  end
  visorFuncEasyPick_b634ba()
  # end: URCap Program Node
  $ 1699 "MoveJ"
  $ 1700 "Waypoint_95" "breakAfter"
  movej(get_inverse_kin(Waypoint_95_p, qnear=Waypoint_95_q), a=1.3962634015954636, v=1.0471975511965976)
  $ 1701 "Wait: 2.0"
  sleep(2.0)
  elif (7 == switch_1):
    $ 1702 "Case 7"
  elif (8 == switch_1):
    $ 1731 "Case 8"
  elif (11 == switch_1):
    $ 1764 "Case 11"
  elif (12 == switch_1):
    $ 1801 "Case 12"
  elif (15 == switch_1):
    $ 1852 "Case 15"
  elif (30 == switch_1):
    $ 1855 "Case 30"
  elif (31 == switch_1):
    $ 1888 "Case 31"
  elif (32 == switch_1):
    $ 1900 "Case 32"
  elif (33 == switch_1):
    $ 1941 "Case 33"
  elif (35 == switch_1):
    $ 2007 "Case 35"
    $ 2008 "Pick the powder container"
    # begin: URCap Program Node
    #   Source: SensoPart VISOR Robotic, 2.0.0, SensoPart Industriesensorik GmbH
    #   Type: VISOR Robotic App
    $ 2011 "VISOR Easy Pick"
    def visorFuncEasyPick_ceefd3():
      # begin: URCap Program Node
      #   Source: SensoPart VISOR Robotic, 2.0.0, SensoPart Industriesensorik GmbH
      #   Type: Easy Pick Setup
      $ 2012 "# 1 Setup" "noBreak"
      local easyPickVisorId = 1
      local easyPickArmMounted = True
      local easyPickSetJob = True
      local easyPickJobName = "Container"
      local easyPickAtImgAcq = False
      local easyPickImgAcqPose = cont_img_pose
      # end: URCap Program Node
      # begin: URCap Program Node
      #   Source: SensoPart VISOR Robotic, 2.0.0, SensoPart Industriesensorik GmbH
      #   Type: Process
      $ 2013 "Process" "noBreak"
      local easyPickObjTaken = False
      local easyPickTrigger = False
      local easyPickPoseIdx = 0
      local easyPickPose = p[0,0,0,0,0,0]
      def easyPickFuncTrigger(visorId, setJob, jobName, arm):
      if (setJob):
        visor_changeJob(visorId, jobName, 6000)
      end
      if (arm):
        visor_trigger(visorId, 6000, "arm")
      else:
        visor_trigger(visorId, 6000)
      end
      global easyPickParts=visor_partsFound(visorId)
      visor_easyPickUpdate(visorId, "parts", visor_partsFound(visorId))
      return visor_getPose3d(visorId, 0)
    end
    while (not easyPickObjTaken):
      easyPickTrigger = (easyPickCount >= visor_partsFound(easyPickVisorId)) or (easyPickCount > 9) or (not visor_easyPickCheckIdent("bb1e48", easyPickVisorId))
      if (easyPickTrigger):
        easyPickCount = 0
      end
      easyPickPoseIdx = easyPickCount
      easyPickPose = visor_getPose3d(easyPickVisorId, easyPickPoseIdx)
      visor_easyPickUpdate(easyPickVisorId, "counter", easyPickPoseIdx)
      # begin: URCap Program Node
      #   Source: SensoPart VISOR Robotic, 2.0.0, SensoPart Industriesensorik GmbH
      #   Type: Image Acquisition Pose
      $ 2014 "Image Acquisition Pose" "noBreak"
      if (easyPickTrigger):
        if (not easyPickAtImgAcq):
          movej(pose_trans(easyPickImgAcqPose,p[0.0000,0.0000,-0.0000,0.0000,0.0000,0.0000]),a=1.3963,v=1.0472,t=0.000000,r=0.000000)
          easyPickAtImgAcq = True
        end
        easyPickPose = easyPickFuncTrigger(easyPickVisorId, easyPickSetJob, easyPickJobName, easyPickArmMounted)
      end
      # end: URCap Program Node
      # begin: URCap Program Node
      #   Source: SensoPart VISOR Robotic, 2.0.0, SensoPart Industriesensorik GmbH
      #   Type: Object Detected
      $ 2015 "Object Detected" "noBreak"
      if (visor_partsFound(easyPickVisorId) > 0):
        $ 2016 "Open Gripper" "noBreak"
        # begin: URCap Program Node
        #   Source: Robotiq_Grippers, 1.8.4.4844, Robotiq Inc.
        #   Type: Gripper
        $ 2017 "Gripper Open (1)" "noBreak"
        if not(gripper_connected[0]):
          popup("Gripper 1 must be connected to run this program.", "No connection", False, True, True)
        end
        if not(rq_is_gripper_activated("1")):
          popup("Gripper 1 is not activated. Go to Installation tab > Gripper to activate it and run the program again.", "Not activated", False, True, True)
        end
        rq_set_pos_spd_for(0, 102, 77, "1")
        rq_wait_pos_spe_for_request(0, 102, 77, "1")
        rq_go_to("1")
        rq_wait("1")
        # end: URCap Program Node
        $ 2018 "MoveJ" "noBreak"
        $ 2019 "Waypoint_13" "noBreak"
        movej(get_inverse_kin(Waypoint_13_p, qnear=Waypoint_13_q), a=1.3962634015954636, v=1.0471975511965976)
        # begin: URCap Program Node
        #   Source: SensoPart VISOR Robotic, 2.0.0, SensoPart Industriesensorik GmbH
        #   Type: Approach Pose
        $ 2020 "Approach Pose" "noBreak"
        movej(pose_trans(easyPickPose,p[0.0000,0.0000,0.0500,0.0000,0.0000,0.0000]),a=1.3963,v=1.0472,t=0.000000,r=0.000000)
        # end: URCap Program Node
        # begin: URCap Program Node
        #   Source: SensoPart VISOR Robotic, 2.0.0, SensoPart Industriesensorik GmbH
        #   Type: Target Pose
        $ 2021 "Target Pose" "noBreak"
        movel(pose_trans(easyPickPose,p[0.0000,0.0000,-0.0000,0.0000,0.0000,0.0000]),a=0.5000,v=0.2500,t=0.000000,r=0.000000)
        # end: URCap Program Node
        $ 2022 "Close Gripper" "noBreak"
        # begin: URCap Program Node
        #   Source: Robotiq_Grippers, 1.8.4.4844, Robotiq Inc.
        #   Type: Gripper
        $ 2023 "Gripper Close (1)" "noBreak"
        if not(gripper_connected[0]):
          popup("Gripper 1 must be connected to run this program.", "No connection", False, True, True)
        end
        if not(rq_is_gripper_activated("1")):
          popup("Gripper 1 is not activated. Go to Installation tab > Gripper to activate it and run the program again.", "Not activated", False, True, True)
        end
        rq_set_pos_spd_for(255, 102, 77, "1")
        rq_wait_pos_spe_for_request(255, 102, 77, "1")
        rq_go_to("1")
        rq_wait("1")
        # end: URCap Program Node
        # begin: URCap Program Node
        #   Source: SensoPart VISOR Robotic, 2.0.0, SensoPart Industriesensorik GmbH
        #   Type: Exit Pose
        $ 2024 "Exit Pose" "noBreak"
        movel(pose_trans(easyPickPose,p[0.0000,0.0000,0.0500,0.0000,0.0000,0.0000]),a=0.5000,v=0.2500,t=0.000000,r=0.000000)
        # end: URCap Program Node
        easyPickObjTaken = True
      end
      # end: URCap Program Node
      # begin: URCap Program Node
      #   Source: SensoPart VISOR Robotic, 2.0.0, SensoPart Industriesensorik GmbH
      #   Type: No Object Detected
      $ 2025 "No Object Detected" "noBreak"
      if (visor_partsFound(easyPickVisorId) < 1):
        $ 2026 "Popup: No Container detected" "noBreak"
        popup("No Container detected", "Message", False, False, blocking=True)
        else:
      end
      # end: URCap Program Node
    end
    easyPickCount = easyPickCount + 1
    visor_easyPickUpdate(easyPickVisorId, "counter", easyPickCount)
    visor_easyPickSetIdent("bb1e48", easyPickVisorId)
    # end: URCap Program Node
  end
  visorFuncEasyPick_ceefd3()
  # end: URCap Program Node
  $ 2027 "MoveJ"
  $ 2029 "Waypoint_70" "breakAfter"
  movej(get_inverse_kin(Waypoint_70_p, qnear=Waypoint_70_q), a=0.6981317007977318, v=0.5235987755982988)
  $ 2030 "Waypoint_2" "breakAfter"
  movej(get_inverse_kin(Waypoint_2_p, qnear=Waypoint_2_q), a=0.8726646259971648, v=0.5235987755982988, r=0.05)
  $ 2031 "Waypoint_3" "breakAfter"
  movej(get_inverse_kin(Waypoint_3_p, qnear=Waypoint_3_q), a=0.6981317007977318, v=0.5235987755982988, r=0.05)
  $ 2032 "MoveL"
  $ 2033 "Waypoint_15" "breakAfter"
  movel(Waypoint_15_p, a=0.5, v=0.1, r=0.05)
  $ 2034 "Waypoint_14" "breakAfter"
  movel(Waypoint_14_p, a=0.3, v=0.1)
  $ 2035 "Waypoint_4" "breakAfter"
  movel(Waypoint_4_p, a=0.3, v=0.05)
  # begin: URCap Program Node
  #   Source: Robotiq_Grippers, 1.8.4.4844, Robotiq Inc.
  #   Type: Gripper
  $ 2036 "Gripper Open (1)"
  if not(gripper_connected[0]):
    popup("Gripper 1 must be connected to run this program.", "No connection", False, True, True)
  end
  if not(rq_is_gripper_activated("1")):
    popup("Gripper 1 is not activated. Go to Installation tab > Gripper to activate it and run the program again.", "Not activated", False, True, True)
  end
  rq_set_pos_spd_for(0, 102, 77, "1")
  rq_wait_pos_spe_for_request(0, 102, 77, "1")
  rq_go_to("1")
  rq_wait("1")
  # end: URCap Program Node
  $ 2037 "MoveL"
  $ 2038 "Waypoint_25" "breakAfter"
  movel(Waypoint_25_p, a=0.3, v=0.1)
  $ 2039 "Waypoint_15" "breakAfter"
  movel(Waypoint_15_p, a=0.5, v=0.1, r=0.05)
  $ 2040 "Home (Safe)"
  movej([-1.2302089344500047, -1.2969853503591224, -1.875639182904262, -1.539621866126728, 1.5731943360401213, -2.80099559440227], a=1.3962634015954636, v=1.0471975511965976)
  elif (36 == switch_1):
    $ 2070 "Case 36"
    $ 2074 "Decap"
    $ 2112 "MoveJ"
    $ 2113 "Waypoint_39" "breakAfter"
    movej(get_inverse_kin(Waypoint_39_p, qnear=Waypoint_39_q), a=1.3962634015954636, v=1.0471975511965976)
    $ 2114 "MoveL"
    $ 2115 "Waypoint_41" "breakAfter"
    movel(Waypoint_41_p, a=0.5, v=0.1)
    $ 2116 "Waypoint_40" "breakAfter"
    movel(Waypoint_40_p, a=0.3, v=0.05)
    # begin: URCap Program Node
    #   Source: Robotiq_Grippers, 1.8.4.4844, Robotiq Inc.
    #   Type: Gripper
    $ 2117 "Gripper Close (1)"
    if not(gripper_connected[0]):
      popup("Gripper 1 must be connected to run this program.", "No connection", False, True, True)
    end
    if not(rq_is_gripper_activated("1")):
      popup("Gripper 1 is not activated. Go to Installation tab > Gripper to activate it and run the program again.", "Not activated", False, True, True)
    end
    rq_set_pos_spd_for(255, 77, 51, "1")
    rq_wait_pos_spe_for_request(255, 77, 51, "1")
    rq_go_to("1")
    rq_wait("1")
    # end: URCap Program Node
    $ 2118 "Loop 2 times"
    Loop_2 = 0
    while (Loop_2 < 2):
      $ 2119 "MoveL"
      $ 2120 "Waypoint_42" "breakAfter"
      movel(Waypoint_42_p, a=1.2, v=0.5)
      $ 2121 "Waypoint_43" "breakAfter"
      movel(Waypoint_43_p, a=1.2, v=0.25)
      # begin: URCap Program Node
      #   Source: Robotiq_Grippers, 1.8.4.4844, Robotiq Inc.
      #   Type: Gripper
      $ 2122 "Gripper Move40mm (1)"
      if not(gripper_connected[0]):
        popup("Gripper 1 must be connected to run this program.", "No connection", False, True, True)
      end
      if not(rq_is_gripper_activated("1")):
        popup("Gripper 1 is not activated. Go to Installation tab > Gripper to activate it and run the program again.", "Not activated", False, True, True)
      end
      rq_set_pos_spd_for(63, 77, 51, "1")
      rq_wait_pos_spe_for_request(63, 77, 51, "1")
      rq_go_to("1")
      rq_wait("1")
      # end: URCap Program Node
      $ 2123 "MoveL"
      $ 2124 "Waypoint_44" "breakAfter"
      movel(Waypoint_44_p, a=1.2, v=0.5)
      $ 2125 "Waypoint_45" "breakAfter"
      movel(Waypoint_45_p, a=1.2, v=0.25)
      # begin: URCap Program Node
      #   Source: Robotiq_Grippers, 1.8.4.4844, Robotiq Inc.
      #   Type: Gripper
      $ 2126 "Gripper Move11mm (1)"
      if not(gripper_connected[0]):
        popup("Gripper 1 must be connected to run this program.", "No connection", False, True, True)
      end
      if not(rq_is_gripper_activated("1")):
        popup("Gripper 1 is not activated. Go to Installation tab > Gripper to activate it and run the program again.", "Not activated", False, True, True)
      end
      rq_set_pos_spd_for(200, 77, 51, "1")
      rq_wait_pos_spe_for_request(200, 77, 51, "1")
      rq_go_to("1")
      rq_wait("1")
      # end: URCap Program Node
      Loop_2 = Loop_2 + 1
    end
    $ 2127 "MoveL"
    $ 2128 "Waypoint_46" "breakAfter"
    movel(Waypoint_46_p, a=0.3, v=0.05)
    $ 2129 "Waypoint_47" "breakAfter"
    movel(Waypoint_47_p, a=0.5, v=0.1)
    $ 2130 "Waypoint_48" "breakAfter"
    movel(Waypoint_48_p, a=1.2, v=0.25)
    $ 2131 "Waypoint_49" "breakAfter"
    movel(Waypoint_49_p, a=1.2, v=0.25)
    # begin: URCap Program Node
    #   Source: Robotiq_Grippers, 1.8.4.4844, Robotiq Inc.
    #   Type: Gripper
    $ 2132 "Gripper Move35mm (1)"
    if not(gripper_connected[0]):
      popup("Gripper 1 must be connected to run this program.", "No connection", False, True, True)
    end
    if not(rq_is_gripper_activated("1")):
      popup("Gripper 1 is not activated. Go to Installation tab > Gripper to activate it and run the program again.", "Not activated", False, True, True)
    end
    rq_set_pos_spd_for(87, 77, 51, "1")
    rq_wait_pos_spe_for_request(87, 77, 51, "1")
    rq_go_to("1")
    rq_wait("1")
    # end: URCap Program Node
    $ 2133 "MoveL"
    $ 2134 "Waypoint_50" "breakAfter"
    movel(Waypoint_50_p, a=1.2, v=0.25)
    $ 2135 "Home (Safe)"
    movej([-1.2302089344500047, -1.2969853503591224, -1.875639182904262, -1.539621866126728, 1.5731943360401213, -2.80099559440227], a=1.3962634015954636, v=1.0471975511965976)
  elif (37 == switch_1):
    $ 2136 "Case 37"
    $ 2137 "Powder dispensing"
    $ 2138 "zero_scale()"
    zero_scale()
    # begin: URCap Program Node
    #   Source: SensoPart VISOR Robotic, 2.0.0, SensoPart Industriesensorik GmbH
    #   Type: VISOR Robotic App
    $ 2139 "VISOR Easy Pick"
    def visorFuncEasyPick_f697d2():
      # begin: URCap Program Node
      #   Source: SensoPart VISOR Robotic, 2.0.0, SensoPart Industriesensorik GmbH
      #   Type: Easy Pick Setup
      $ 2140 "# 1 Setup" "noBreak"
      local easyPickVisorId = 1
      local easyPickArmMounted = True
      local easyPickSetJob = True
      local easyPickJobName = "Weigh_scale"
      local easyPickAtImgAcq = False
      local easyPickImgAcqPose = cont_img_pose
      # end: URCap Program Node
      # begin: URCap Program Node
      #   Source: SensoPart VISOR Robotic, 2.0.0, SensoPart Industriesensorik GmbH
      #   Type: Process
      $ 2141 "Process" "noBreak"
      local easyPickObjTaken = False
      local easyPickTrigger = False
      local easyPickPoseIdx = 0
      local easyPickPose = p[0,0,0,0,0,0]
      def easyPickFuncTrigger(visorId, setJob, jobName, arm):
      if (setJob):
        visor_changeJob(visorId, jobName, 6000)
      end
      if (arm):
        visor_trigger(visorId, 6000, "arm")
      else:
        visor_trigger(visorId, 6000)
      end
      global easyPickParts_4=visor_partsFound(visorId)
      visor_easyPickUpdate(visorId, "parts", visor_partsFound(visorId))
      return visor_getPose3d(visorId, 0)
    end
    while (not easyPickObjTaken):
      easyPickTrigger = (easyPickCount_4 >= visor_partsFound(easyPickVisorId)) or (easyPickCount_4 > 9) or (not visor_easyPickCheckIdent("db3fd8", easyPickVisorId))
      if (easyPickTrigger):
        easyPickCount_4 = 0
      end
      easyPickPoseIdx = easyPickCount_4
      easyPickPose = visor_getPose3d(easyPickVisorId, easyPickPoseIdx)
      visor_easyPickUpdate(easyPickVisorId, "counter", easyPickPoseIdx)
      # begin: URCap Program Node
      #   Source: SensoPart VISOR Robotic, 2.0.0, SensoPart Industriesensorik GmbH
      #   Type: Image Acquisition Pose
      $ 2142 "Image Acquisition Pose" "noBreak"
      if (easyPickTrigger):
        if (not easyPickAtImgAcq):
          movej(pose_trans(easyPickImgAcqPose,p[0.0000,0.0000,-0.0000,0.0000,0.0000,0.0000]),a=1.3963,v=1.0472,t=0.000000,r=0.000000)
          easyPickAtImgAcq = True
        end
        easyPickPose = easyPickFuncTrigger(easyPickVisorId, easyPickSetJob, easyPickJobName, easyPickArmMounted)
      end
      # end: URCap Program Node
      # begin: URCap Program Node
      #   Source: SensoPart VISOR Robotic, 2.0.0, SensoPart Industriesensorik GmbH
      #   Type: Object Detected
      $ 2143 "Object Detected" "noBreak"
      if (visor_partsFound(easyPickVisorId) > 0):
        $ 2144 "Open Gripper" "noBreak"
        $ 2145 "MoveL" "noBreak"
        $ 2146 "Weight_value≔get_weight()" "noBreak"
        global Weight_value=get_weight()
        # begin: URCap Program Node
        #   Source: Robotiq_Grippers, 1.8.4.4844, Robotiq Inc.
        #   Type: Gripper
        $ 2147 "Gripper Open (1)" "noBreak"
        if not(gripper_connected[0]):
          popup("Gripper 1 must be connected to run this program.", "No connection", False, True, True)
        end
        if not(rq_is_gripper_activated("1")):
          popup("Gripper 1 is not activated. Go to Installation tab > Gripper to activate it and run the program again.", "Not activated", False, True, True)
        end
        rq_set_pos_spd_for(0, 77, 77, "1")
        rq_wait_pos_spe_for_request(0, 77, 77, "1")
        rq_go_to("1")
        rq_wait("1")
        # end: URCap Program Node
        $ 2148 "Waypoint_53" "noBreak"
        movel(Waypoint_53_p, a=0.6, v=0.15, r=0.05)
        $ 2149 "Spatula_above" "noBreak"
        movel(Spatula_above_p, a=0.6, v=0.15)
        $ 2150 "Spatula_pick" "noBreak"
        movel(Spatula_pick_p, a=0.6, v=0.15)
        # begin: URCap Program Node
        #   Source: Robotiq_Grippers, 1.8.4.4844, Robotiq Inc.
        #   Type: Gripper
        $ 2151 "Gripper Close (1)" "noBreak"
        if not(gripper_connected[0]):
          popup("Gripper 1 must be connected to run this program.", "No connection", False, True, True)
        end
        if not(rq_is_gripper_activated("1")):
          popup("Gripper 1 is not activated. Go to Installation tab > Gripper to activate it and run the program again.", "Not activated", False, True, True)
        end
        rq_set_pos_spd_for(255, 77, 77, "1")
        rq_wait_pos_spe_for_request(255, 77, 77, "1")
        rq_go_to("1")
        rq_wait("1")
        # end: URCap Program Node
        $ 2152 "Spatula_above" "noBreak"
        movel(Spatula_above_p, a=0.6, v=0.15)
        $ 2153 "Popup: Connect the vibration motor" "noBreak"
        popup("Connect the vibration motor", "Message", False, False, blocking=True)
        $ 2154 "tare_scale()" "noBreak"
        tare_scale()
        $ 2155 "container_start" "noBreak"
        movel(container_start_p, a=0.3, v=0.1)
        $ 2156 "container_wp_1" "noBreak"
        movel(container_wp_1_p, a=0.3, v=0.05)
        $ 2157 "Loop 1 times" "noBreak"
        Loop_9 = 0
        while (Loop_9 < 1):
          $ 2158 "Waypoint_55" "noBreak"
          global move_thread_flag_2158=0
          thread move_thread_2158():
            enter_critical
            move_thread_flag_2158 = 1
            movel(Waypoint_55_p, a=0.5, v=0.07)
            move_thread_flag_2158 = 2
            exit_critical
          end
          move_thread_flag_2158 = 0
          move_thread_han_2158 = run move_thread_2158()
          while (True):
            sleep(1.0E-10)
            if (move_thread_flag_2158 > 1):
              join move_thread_han_2158
              break
            end
            sync()
          end
          $ 2160 "Waypoint_56" "noBreak"
          movel(Waypoint_56_p, a=0.3, v=0.05)
          $ 2161 "Waypoint_74" "noBreak"
          movel(Waypoint_74_p, a=0.6, v=0.15)
          $ 2162 "Set AO[0]=3.0" "noBreak"
          set_standard_analog_out(0, 0.3)
          $ 2163 "Wait: 2.0" "noBreak"
          sleep(2.0)
          $ 2164 "Set AO[0]=0.0" "noBreak"
          set_standard_analog_out(0, 0.0)
          Loop_9 = Loop_9 + 1
        end
        $ 2168 "ftr_scoop2" "noBreak"
        movel(ftr_scoop2_p, a=0.3, v=0.05)
        $ 2169 "aftr_scoo3" "noBreak"
        movel(aftr_scoo3_p, a=0.3, v=0.05)
        $ 2170 "MoveJ" "noBreak"
        $ 2171 "Waypoint_60" "noBreak"
        movej(get_inverse_kin(Waypoint_60_p, qnear=Waypoint_60_q), a=0.5235987755982988, v=0.3490658503988659, r=0.05)
        $ 2172 "Waypoint_61" "noBreak"
        movej(get_inverse_kin(Waypoint_61_p, qnear=Waypoint_61_q), a=0.5235987755982988, v=0.3490658503988659, r=0.05)
        # begin: URCap Program Node
        #   Source: SensoPart VISOR Robotic, 2.0.0, SensoPart Industriesensorik GmbH
        #   Type: Approach Pose
        $ 2173 "Approach Pose" "noBreak"
        movej(pose_trans(easyPickPose,p[0.0000,0.0000,0.0500,0.0000,0.0000,0.0000]),a=0.4363,v=0.3491,t=0.000000,r=0.000000)
        # end: URCap Program Node
        # begin: URCap Program Node
        #   Source: SensoPart VISOR Robotic, 2.0.0, SensoPart Industriesensorik GmbH
        #   Type: Target Pose
        $ 2174 "Target Pose" "noBreak"
        movel(pose_trans(easyPickPose,p[0.0000,0.0000,-0.0000,0.0000,0.0000,0.0000]),a=0.1000,v=0.0500,t=0.000000,r=0.000000)
        # end: URCap Program Node
        $ 2175 "Close Gripper" "noBreak"
        $ 2176 "dispense_pos≔get_actual_tcp_pose()" "noBreak"
        global dispense_pos= get_actual_tcp_pose ()
        $ 2177 "MoveL" "noBreak"
        $ 2178 "Start_thread≔ True " "noBreak"
        global Start_thread=  True
        $ 2179 "vib_mot_thread≔ True " "noBreak"
        global vib_mot_thread=  True
        $ 2180 "tilt_angle≔current_pose[4]" "noBreak"
        global tilt_angle=current_pose[4]
        $ 2181 "Wait: 0.5" "noBreak"
        sleep(0.5)
        $ 2182 "Loop Weight_value≤Target_weight and tilt_angle≤-0.40" "noBreak"
        thread Thread_while_2182():
          while (True):
            $ 2183 "current_error≔Target_weight-Weight_value" "noBreak"
            global current_error=Target_weight-Weight_value
            $ 2184 "Integral_error≔Integral_error+current_error*dt" "noBreak"
            global Integral_error=Integral_error+current_error*dt
            $ 2185 "derivative≔(current_error-previous_error)/dt" "noBreak"
            global derivative=(current_error-previous_error)/dt
            $ 2186 "tilt_increment≔(kp*current_error)+(ki*Integral_error)+(kd*derivative)" "noBreak"
            global tilt_increment=(kp*current_error)+(ki*Integral_error)+(kd*derivative)
            $ 2187 "current_pose≔get_actual_tcp_pose()" "noBreak"
            global current_pose= get_actual_tcp_pose ()
            $ 2188 "tilt_angle≔current_pose[4]" "noBreak"
            global tilt_angle=current_pose[4]
            $ 2189 "tilt_pose≔pose_trans(current_pose, p[(tilt_increment/7), 0, 0, 0, tilt_increment, 0])" "noBreak"
            global tilt_pose=pose_trans(current_pose, p[(tilt_increment/7), 0, 0, 0, tilt_increment, 0])
            $ 2190 "movel(tilt_pose, a=0.025, v=0.015, r=0.00001)" "noBreak"
            movel(tilt_pose, a=0.025, v=0.015, r=0.00001)
            $ 2191 "previous_error≔current_error" "noBreak"
            global previous_error=current_error
          end
        end
        if (Weight_value <= Target_weight  and  tilt_angle <= -0.40):
          global thread_handler_2182=run Thread_while_2182()
          while (Weight_value <= Target_weight  and  tilt_angle <= -0.40):
            sync()
          end
          kill thread_handler_2182
        end
        $ 2192 "Start_thread≔ False " "noBreak"
        global Start_thread=  False
        $ 2194 "Weight_value≔get_weight()" "noBreak"
        global Weight_value=get_weight()
        $ 2195 "tilt_angle≔-1" "noBreak"
        global tilt_angle=-1
        $ 2196 "Wait: 0.5" "noBreak"
        sleep(0.5)
        $ 2197 "vib_mot_thread≔ False " "noBreak"
        global vib_mot_thread=  False
        $ 2198 "MoveL" "noBreak"
        $ 2199 "dispense_pos" "noBreak"
        movel(dispense_pos, a=0.2, v=0.05)
        $ 2200 "Integral_error≔0" "noBreak"
        global Integral_error=0
        $ 2201 "current_error≔0" "noBreak"
        global current_error=0
        $ 2202 "previous_error≔0" "noBreak"
        global previous_error=0
        $ 2203 "Set AO[0]=0.0" "noBreak"
        set_standard_analog_out(0, 0.0)
        # begin: URCap Program Node
        #   Source: SensoPart VISOR Robotic, 2.0.0, SensoPart Industriesensorik GmbH
        #   Type: Exit Pose
        $ 2204 "Exit Pose" "noBreak"
        movel(pose_trans(easyPickPose,p[0.0000,0.0000,-0.0000,0.0000,0.0000,0.0000]),a=0.5000,v=0.2500,t=0.000000,r=0.000000)
        # end: URCap Program Node
        easyPickObjTaken = True
      end
      # end: URCap Program Node
      # begin: URCap Program Node
      #   Source: SensoPart VISOR Robotic, 2.0.0, SensoPart Industriesensorik GmbH
      #   Type: No Object Detected
      $ 2205 "No Object Detected" "noBreak"
      if (visor_partsFound(easyPickVisorId) < 1):
        $ 2206 "Popup: No weigh scale detected" "noBreak"
        popup("No weigh scale detected", "Message", False, False, blocking=True)
        else:
      end
      # end: URCap Program Node
    end
    easyPickCount_4 = easyPickCount_4 + 1
    visor_easyPickUpdate(easyPickVisorId, "counter", easyPickCount_4)
    visor_easyPickSetIdent("db3fd8", easyPickVisorId)
    # end: URCap Program Node
  end
  visorFuncEasyPick_f697d2()
  # end: URCap Program Node
  $ 2207 "powder dispensing"
  $ 2209 "Loop Weight_value<Target_weight"
  while (Weight_value<Target_weight):
    $ 2210 "MoveL"
    $ 2211 "Waypoint_75" "breakAfter"
    movel(Waypoint_75_p, a=0.3, v=0.05, r=0.05)
    $ 2212 "ftr_scoop2" "breakAfter"
    movel(ftr_scoop2_p, a=0.3, v=0.05)
    $ 2213 "aftr_scoop1" "breakAfter"
    movel(aftr_scoop1_p, a=0.3, v=0.05)
    $ 2214 "After_disp_3" "breakAfter"
    movel(After_disp_3_p, a=0.3, v=0.05)
    $ 2215 "Loop 1 times"
    Loop_13 = 0
    while (Loop_13 < 1):
      $ 2216 "Waypoint_55" "breakAfter"
      global move_thread_flag_2216=0
      thread move_thread_2216():
        enter_critical
        move_thread_flag_2216 = 1
        movel(Waypoint_55_p, a=0.5, v=0.07)
        move_thread_flag_2216 = 2
        exit_critical
      end
      move_thread_flag_2216 = 0
      move_thread_han_2216 = run move_thread_2216()
      while (True):
        sleep(1.0E-10)
        if (move_thread_flag_2216 > 1):
          join move_thread_han_2216
          break
        end
        sync()
      end
      $ 2218 "Waypoint_56" "breakAfter"
      movel(Waypoint_56_p, a=0.3, v=0.05)
      $ 2219 "Waypoint_74" "breakAfter"
      movel(Waypoint_74_p, a=0.3, v=0.05)
      $ 2220 "Set AO[0]=3.0"
      set_standard_analog_out(0, 0.3)
      $ 2221 "Wait: 2.0"
      sleep(2.0)
      $ 2222 "Set AO[0]=0.0"
      set_standard_analog_out(0, 0.0)
      Loop_13 = Loop_13 + 1
    end
    $ 2223 "ftr_scoop2" "breakAfter"
    movel(ftr_scoop2_p, a=0.3, v=0.05)
    $ 2224 "aftr_scoo3" "breakAfter"
    movel(aftr_scoo3_p, a=0.3, v=0.05)
    $ 2225 "MoveJ"
    $ 2226 "Waypoint_60" "breakAfter"
    movej(get_inverse_kin(Waypoint_60_p, qnear=Waypoint_60_q), a=0.5235987755982988, v=0.3490658503988659, r=0.05)
    $ 2227 "Waypoint_61" "breakAfter"
    movej(get_inverse_kin(Waypoint_61_p, qnear=Waypoint_61_q), a=0.5235987755982988, v=0.3490658503988659, r=0.05)
    $ 2228 "Waypoint_62" "breakAfter"
    movej(get_inverse_kin(Waypoint_62_p, qnear=Waypoint_62_q), a=0.5235987755982988, v=0.3490658503988659)
    $ 2229 "MoveL"
    $ 2230 "Start_thread≔ True "
    global Start_thread=  True
    $ 2231 "dispense_pos" "breakAfter"
    movel(dispense_pos, a=0.2, v=0.05)
    $ 2232 "vib_mot_thread≔ True "
    global vib_mot_thread=  True
    $ 2233 "Wait: 0.5"
    sleep(0.5)
    $ 2234 "Loop Weight_value≤Target_weight and tilt_angle≤-0.40"
    thread Thread_while_2234():
      while (True):
        $ 2235 "current_error≔Target_weight-Weight_value"
        global current_error=Target_weight-Weight_value
        $ 2236 "Integral_error≔Integral_error+current_error*dt"
        global Integral_error=Integral_error+current_error*dt
        $ 2237 "derivative≔(current_error-previous_error)/dt"
        global derivative=(current_error-previous_error)/dt
        $ 2238 "tilt_increment≔(kp*current_error)+(ki*Integral_error)+(kd*derivative)"
        global tilt_increment=(kp*current_error)+(ki*Integral_error)+(kd*derivative)
        $ 2239 "current_pose≔get_actual_tcp_pose()"
        global current_pose= get_actual_tcp_pose ()
        $ 2240 "tilt_angle≔current_pose[4]"
        global tilt_angle=current_pose[4]
        $ 2241 "tilt_pose≔pose_trans(current_pose, p[(tilt_increment/7), 0, 0, 0, tilt_increment, 0])"
        global tilt_pose=pose_trans(current_pose, p[(tilt_increment/7), 0, 0, 0, tilt_increment, 0])
        $ 2242 "movel(tilt_pose, a=0.025, v=0.015, r=0.00001)"
        movel(tilt_pose, a=0.025, v=0.015, r=0.00001)
        $ 2243 "previous_error≔current_error"
        global previous_error=current_error
        $ 2244 "Wait: 0.01"
        sleep(0.01)
      end
    end
    if (Weight_value <= Target_weight  and  tilt_angle <= -0.40):
      global thread_handler_2234=run Thread_while_2234()
      while (Weight_value <= Target_weight  and  tilt_angle <= -0.40):
        sync()
      end
      kill thread_handler_2234
    end
    $ 2245 "Start_thread≔ False "
    global Start_thread=  False
    $ 2246 "Set AO[0]=0.0"
    set_standard_analog_out(0, 0.0)
    $ 2247 "vib_mot_thread≔ False "
    global vib_mot_thread=  False
    $ 2249 "Weight_value≔get_weight()"
    global Weight_value=get_weight()
    $ 2250 "tilt_angle≔-1"
    global tilt_angle=-1
    $ 2251 "Wait: 0.5"
    sleep(0.5)
    $ 2252 "MoveL"
    $ 2253 "dispense_pos" "breakAfter"
    movel(dispense_pos, a=0.2, v=0.05)
    $ 2254 "Integral_error≔0"
    global Integral_error=0
    $ 2255 "current_error≔0"
    global current_error=0
    $ 2256 "previous_error≔0"
    global previous_error=0
  end
  $ 2257 "MoveL"
  $ 2258 "aftr_scoo3" "breakAfter"
  movel(aftr_scoo3_p, a=0.3, v=0.1)
  $ 2259 "ftr_scoop2" "breakAfter"
  movel(ftr_scoop2_p, a=0.4, v=0.1)
  $ 2260 "aftr_scoop1" "breakAfter"
  movel(aftr_scoop1_p, a=0.4, v=0.1)
  $ 2261 "After_disp_3" "breakAfter"
  movel(After_disp_3_p, a=0.4, v=0.1)
  $ 2262 "Set AO[0]=3.0"
  set_standard_analog_out(0, 0.3)
  $ 2263 "Wait: 2.0"
  sleep(2.0)
  $ 2264 "Set AO[0]=0.0"
  set_standard_analog_out(0, 0.0)
  $ 2265 "aftr_scoop1" "breakAfter"
  movel(aftr_scoop1_p, a=1.2, v=0.25)
  $ 2266 "ftr_scoop2" "breakAfter"
  movel(ftr_scoop2_p, a=0.4, v=0.1)
  $ 2267 "Waypoint_63" "breakAfter"
  movel(Waypoint_63_p, a=1.2, v=0.25, r=0.05)
  $ 2268 "Start" "breakAfter"
  movel(Start_p, a=0.6, v=0.15)
  $ 2269 "Popup: Powder dispensed successfully..."
  popup("Powder dispensed successfully...", "Message", False, False, blocking=True)
  elif (38 == switch_1):
    $ 2270 "Case 38"
    $ 2271 "PowderA(M200)"
    # begin: URCap Program Node
    #   Source: SensoPart VISOR Robotic, 2.0.0, SensoPart Industriesensorik GmbH
    #   Type: VISOR Robotic App
    $ 2272 "VISOR Easy Pick"
    def visorFuncEasyPick_c25fc1():
      # begin: URCap Program Node
      #   Source: SensoPart VISOR Robotic, 2.0.0, SensoPart Industriesensorik GmbH
      #   Type: Easy Pick Setup
      $ 2273 "# 1 Setup" "noBreak"
      local easyPickVisorId = 1
      local easyPickArmMounted = True
      local easyPickSetJob = True
      local easyPickJobName = "PowderA"
      local easyPickAtImgAcq = False
      local easyPickImgAcqPose = cont_img_pose
      # end: URCap Program Node
      # begin: URCap Program Node
      #   Source: SensoPart VISOR Robotic, 2.0.0, SensoPart Industriesensorik GmbH
      #   Type: Process
      $ 2274 "Process" "noBreak"
      local easyPickObjTaken = False
      local easyPickTrigger = False
      local easyPickPoseIdx = 0
      local easyPickPose = p[0,0,0,0,0,0]
      def easyPickFuncTrigger(visorId, setJob, jobName, arm):
      if (setJob):
        visor_changeJob(visorId, jobName, 6000)
      end
      if (arm):
        visor_trigger(visorId, 6000, "arm")
      else:
        visor_trigger(visorId, 6000)
      end
      global easyPickParts_6=visor_partsFound(visorId)
      visor_easyPickUpdate(visorId, "parts", visor_partsFound(visorId))
      return visor_getPose3d(visorId, 0)
    end
    while (not easyPickObjTaken):
      easyPickTrigger = (easyPickCount_6 >= visor_partsFound(easyPickVisorId)) or (easyPickCount_6 > 9) or (not visor_easyPickCheckIdent("617d47", easyPickVisorId))
      if (easyPickTrigger):
        easyPickCount_6 = 0
      end
      easyPickPoseIdx = easyPickCount_6
      easyPickPose = visor_getPose3d(easyPickVisorId, easyPickPoseIdx)
      visor_easyPickUpdate(easyPickVisorId, "counter", easyPickPoseIdx)
      # begin: URCap Program Node
      #   Source: SensoPart VISOR Robotic, 2.0.0, SensoPart Industriesensorik GmbH
      #   Type: Image Acquisition Pose
      $ 2275 "Image Acquisition Pose" "noBreak"
      if (easyPickTrigger):
        if (not easyPickAtImgAcq):
          movej(pose_trans(easyPickImgAcqPose,p[0.0000,0.0000,-0.0000,0.0000,0.0000,0.0000]),a=1.3963,v=1.0472,t=0.000000,r=0.000000)
          easyPickAtImgAcq = True
        end
        easyPickPose = easyPickFuncTrigger(easyPickVisorId, easyPickSetJob, easyPickJobName, easyPickArmMounted)
      end
      # end: URCap Program Node
      # begin: URCap Program Node
      #   Source: SensoPart VISOR Robotic, 2.0.0, SensoPart Industriesensorik GmbH
      #   Type: Object Detected
      $ 2276 "Object Detected" "noBreak"
      if (visor_partsFound(easyPickVisorId) > 0):
        $ 2277 "Open Gripper" "noBreak"
        # begin: URCap Program Node
        #   Source: Robotiq_Grippers, 1.8.4.4844, Robotiq Inc.
        #   Type: Gripper
        $ 2278 "Gripper Open (1)" "noBreak"
        if not(gripper_connected[0]):
          popup("Gripper 1 must be connected to run this program.", "No connection", False, True, True)
        end
        if not(rq_is_gripper_activated("1")):
          popup("Gripper 1 is not activated. Go to Installation tab > Gripper to activate it and run the program again.", "Not activated", False, True, True)
        end
        rq_set_pos_spd_for(0, 77, 77, "1")
        rq_wait_pos_spe_for_request(0, 77, 77, "1")
        rq_go_to("1")
        rq_wait("1")
        # end: URCap Program Node
        $ 2279 "MoveJ" "noBreak"
        $ 2280 "Waypoint_76" "noBreak"
        movej(get_inverse_kin(Waypoint_76_p, qnear=Waypoint_76_q), a=1.3962634015954636, v=1.0471975511965976)
        # begin: URCap Program Node
        #   Source: SensoPart VISOR Robotic, 2.0.0, SensoPart Industriesensorik GmbH
        #   Type: Approach Pose
        $ 2281 "Approach Pose" "noBreak"
        movej(pose_trans(easyPickPose,p[0.0000,0.0000,0.0500,0.0000,0.0000,0.0000]),a=1.3963,v=1.0472,t=0.000000,r=0.000000)
        # end: URCap Program Node
        # begin: URCap Program Node
        #   Source: SensoPart VISOR Robotic, 2.0.0, SensoPart Industriesensorik GmbH
        #   Type: Target Pose
        $ 2282 "Target Pose" "noBreak"
        movel(pose_trans(easyPickPose,p[0.0000,0.0000,-0.0000,0.0000,0.0000,0.0000]),a=0.5000,v=0.2500,t=0.000000,r=0.000000)
        # end: URCap Program Node
        $ 2283 "Close Gripper" "noBreak"
        # begin: URCap Program Node
        #   Source: Robotiq_Grippers, 1.8.4.4844, Robotiq Inc.
        #   Type: Gripper
        $ 2284 "Gripper Move0mm (1)" "noBreak"
        if not(gripper_connected[0]):
          popup("Gripper 1 must be connected to run this program.", "No connection", False, True, True)
        end
        if not(rq_is_gripper_activated("1")):
          popup("Gripper 1 is not activated. Go to Installation tab > Gripper to activate it and run the program again.", "Not activated", False, True, True)
        end
        rq_set_pos_spd_for(247, 77, 77, "1")
        rq_wait_pos_spe_for_request(247, 77, 77, "1")
        rq_go_to("1")
        rq_wait("1")
        # end: URCap Program Node
        # begin: URCap Program Node
        #   Source: SensoPart VISOR Robotic, 2.0.0, SensoPart Industriesensorik GmbH
        #   Type: Exit Pose
        $ 2285 "Exit Pose" "noBreak"
        movel(pose_trans(easyPickPose,p[0.0000,0.0000,0.0500,0.0000,0.0000,0.0000]),a=0.5000,v=0.2500,t=0.000000,r=0.000000)
        # end: URCap Program Node
        easyPickObjTaken = True
      end
      # end: URCap Program Node
      # begin: URCap Program Node
      #   Source: SensoPart VISOR Robotic, 2.0.0, SensoPart Industriesensorik GmbH
      #   Type: No Object Detected
      $ 2286 "No Object Detected" "noBreak"
      if (visor_partsFound(easyPickVisorId) < 1):
        $ 2287 "Popup: No Powder container is detected" "noBreak"
        popup("No Powder container is detected", "Message", False, False, blocking=True)
        else:
      end
      # end: URCap Program Node
    end
    easyPickCount_6 = easyPickCount_6 + 1
    visor_easyPickUpdate(easyPickVisorId, "counter", easyPickCount_6)
    visor_easyPickSetIdent("617d47", easyPickVisorId)
    # end: URCap Program Node
  end
  visorFuncEasyPick_c25fc1()
  # end: URCap Program Node
  $ 2288 "MoveJ"
  $ 2289 "PowderA_wayp1" "breakAfter"
  movej(get_inverse_kin(PowderA_wayp1_p, qnear=PowderA_wayp1_q), a=1.3962634015954636, v=1.0471975511965976, r=0.05)
  $ 2290 "MoveL"
  $ 2291 "Waypoint_80" "breakAfter"
  movel(Waypoint_80_p, a=1.2, v=0.25)
  $ 2292 "MoveL"
  $ 2293 "Decapp_above" "breakAfter"
  movel(Decapp_above_p, a=1.2, v=0.25)
  $ 2294 "Set GRP_3F_Open=On"
  set_standard_digital_out(5, True)
  $ 2295 "Wait: 0.5"
  sleep(0.5)
  $ 2296 "Decapp_place" "breakAfter"
  movel(Decapp_place_p, a=0.3, v=0.05)
  $ 2297 "Set GRP_3F_Open=Off"
  set_standard_digital_out(5, False)
  $ 2298 "Wait: 0.5"
  sleep(0.5)
  # begin: URCap Program Node
  #   Source: Robotiq_Grippers, 1.8.4.4844, Robotiq Inc.
  #   Type: Gripper
  $ 2299 "Gripper Move40mm (1)"
  if not(gripper_connected[0]):
    popup("Gripper 1 must be connected to run this program.", "No connection", False, True, True)
  end
  if not(rq_is_gripper_activated("1")):
    popup("Gripper 1 is not activated. Go to Installation tab > Gripper to activate it and run the program again.", "Not activated", False, True, True)
  end
  rq_set_pos_spd_for(64, 77, 77, "1")
  rq_wait_pos_spe_for_request(64, 77, 77, "1")
  rq_go_to("1")
  rq_wait("1")
  # end: URCap Program Node
  $ 2300 "MoveL"
  $ 2301 "Decapp_above" "breakAfter"
  movel(Decapp_above_p, a=1.2, v=0.25)
  $ 2302 "Waypoint_78" "breakAfter"
  movel(Waypoint_78_p, a=1.2, v=0.25, r=0.05)
  $ 2303 "Home (Safe)"
  movej([-1.2302089344500047, -1.2969853503591224, -1.875639182904262, -1.539621866126728, 1.5731943360401213, -2.80099559440227], a=1.3962634015954636, v=1.0471975511965976)
  elif (39 == switch_1):
    $ 2304 "Case 39"
    $ 2305 "Decap Container A"
    $ 2306 "MoveL"
    $ 2307 "Waypoint_81" "breakAfter"
    movel(Waypoint_81_p, a=1.2, v=0.25)
    $ 2308 "Waypoint_79" "breakAfter"
    movel(Waypoint_79_p, a=1.2, v=0.25)
    # begin: URCap Program Node
    #   Source: Robotiq_Grippers, 1.8.4.4844, Robotiq Inc.
    #   Type: Gripper
    $ 2309 "Gripper Move22mm (1)"
    if not(gripper_connected[0]):
      popup("Gripper 1 must be connected to run this program.", "No connection", False, True, True)
    end
    if not(rq_is_gripper_activated("1")):
      popup("Gripper 1 is not activated. Go to Installation tab > Gripper to activate it and run the program again.", "Not activated", False, True, True)
    end
    rq_set_pos_spd_for(145, 77, 77, "1")
    rq_wait_pos_spe_for_request(145, 77, 77, "1")
    rq_go_to("1")
    rq_wait("1")
    # end: URCap Program Node
    $ 2310 "Decap"
    $ 2311 "Action_Info≔'decapping'"
    global Action_Info="decapping"
    $ 2312 "Set GRP_3F_Enable=On"
    set_standard_digital_out(4, True)
    $ 2313 "Set GRP_3F_Decap=On"
    set_standard_digital_out(3, True)
    $ 2314 "Force"
    sleep(0.02)
    zero_ftsensor()
    force_mode(p[0.0,0.0,0.0,0.0,0.0,0.0], [0, 0, 1, 0, 0, 0], [0.0, 0.0, 2.0, 0.0, 0.0, 0.0], 2, [0.1, 0.1, 5.0E-4, 0.3490658503988659, 0.3490658503988659, 0.3490658503988659])
    $ 2315 "check_decapping(offset=0.010, timeout=4, abort=CMD_Hold)" "noBreak"
    check_decapping(offset=0.010, timeout=4, abort=CMD_Hold)
    end_force_mode()
    stopl(5.0)
    $ 2316 "Set GRP_3F_Decap=Off"
    set_standard_digital_out(3, False)
    $ 2317 "Set GRP_3F_Enable=Off"
    set_standard_digital_out(4, False)
    $ 2318 "MoveL"
    $ 2319 "Waypoint_82" "breakAfter"
    movel(Waypoint_82_p, a=1.2, v=0.25)
    $ 2320 "Cap_above" "breakAfter"
    movel(Cap_above_p, a=1.2, v=0.25, r=0.05)
    $ 2321 "Cap_Place" "breakAfter"
    movel(Cap_Place_p, a=1.2, v=0.25)
    # begin: URCap Program Node
    #   Source: Robotiq_Grippers, 1.8.4.4844, Robotiq Inc.
    #   Type: Gripper
    $ 2322 "Gripper Move39mm (1)"
    if not(gripper_connected[0]):
      popup("Gripper 1 must be connected to run this program.", "No connection", False, True, True)
    end
    if not(rq_is_gripper_activated("1")):
      popup("Gripper 1 is not activated. Go to Installation tab > Gripper to activate it and run the program again.", "Not activated", False, True, True)
    end
    rq_set_pos_spd_for(67, 77, 77, "1")
    rq_wait_pos_spe_for_request(67, 77, 77, "1")
    rq_go_to("1")
    rq_wait("1")
    # end: URCap Program Node
    $ 2323 "Cap_above" "breakAfter"
    movel(Cap_above_p, a=1.2, v=0.25)
    $ 2324 "Home (Safe)"
    movej([-1.2302089344500047, -1.2969853503591224, -1.875639182904262, -1.539621866126728, 1.5731943360401213, -2.80099559440227], a=1.3962634015954636, v=1.0471975511965976)
    $ 2325 "Placing container in th tilt station (Platform version)"
    # begin: URCap Program Node
    #   Source: Robotiq_Grippers, 1.8.4.4844, Robotiq Inc.
    #   Type: Gripper
    $ 2326 "Gripper Open (1)"
    if not(gripper_connected[0]):
      popup("Gripper 1 must be connected to run this program.", "No connection", False, True, True)
    end
    if not(rq_is_gripper_activated("1")):
      popup("Gripper 1 is not activated. Go to Installation tab > Gripper to activate it and run the program again.", "Not activated", False, True, True)
    end
    rq_set_pos_spd_for(0, 77, 77, "1")
    rq_wait_pos_spe_for_request(0, 77, 77, "1")
    rq_go_to("1")
    rq_wait("1")
    # end: URCap Program Node
    $ 2327 "MoveL"
    $ 2328 "OP_PowderA2" "breakAfter"
    movel(OP_PowderA2_p, a=1.2, v=0.25)
    $ 2329 "OP_PowderA_abov" "breakAfter"
    movel(OP_PowderA_abov_p, a=1.2, v=0.25)
    $ 2330 "OP_PowderA_pick" "breakAfter"
    movel(OP_PowderA_pick_p, a=1.2, v=0.25)
    # begin: URCap Program Node
    #   Source: Robotiq_Grippers, 1.8.4.4844, Robotiq Inc.
    #   Type: Gripper
    $ 2331 "Gripper Close (1)"
    if not(gripper_connected[0]):
      popup("Gripper 1 must be connected to run this program.", "No connection", False, True, True)
    end
    if not(rq_is_gripper_activated("1")):
      popup("Gripper 1 is not activated. Go to Installation tab > Gripper to activate it and run the program again.", "Not activated", False, True, True)
    end
    rq_set_pos_spd_for(255, 77, 77, "1")
    rq_wait_pos_spe_for_request(255, 77, 77, "1")
    rq_go_to("1")
    rq_wait("1")
    # end: URCap Program Node
    $ 2332 "Wait: 0.5"
    sleep(0.5)
    $ 2333 "Set GRP_3F_Open=On"
    set_standard_digital_out(5, True)
    $ 2334 "OP_PowderA_abov" "breakAfter"
    movel(OP_PowderA_abov_p, a=0.3, v=0.05)
    $ 2335 "Tilt_above" "breakAfter"
    movel(Tilt_above_p, a=1.2, v=0.25)
    $ 2336 "Tilt_place" "breakAfter"
    movel(Tilt_place_p, a=0.3, v=0.05)
    # begin: URCap Program Node
    #   Source: Robotiq_Grippers, 1.8.4.4844, Robotiq Inc.
    #   Type: Gripper
    $ 2337 "Gripper Open (1)"
    if not(gripper_connected[0]):
      popup("Gripper 1 must be connected to run this program.", "No connection", False, True, True)
    end
    if not(rq_is_gripper_activated("1")):
      popup("Gripper 1 is not activated. Go to Installation tab > Gripper to activate it and run the program again.", "Not activated", False, True, True)
    end
    rq_set_pos_spd_for(0, 77, 77, "1")
    rq_wait_pos_spe_for_request(0, 77, 77, "1")
    rq_go_to("1")
    rq_wait("1")
    # end: URCap Program Node
    $ 2338 "Tilt_above" "breakAfter"
    movel(Tilt_above_p, a=1.2, v=0.25)
    $ 2346 "MoveP"
    $ 2347 "Waypoint_52" "breakAfter"
    movep(Waypoint_52_p, a=0.3, v=0.05, r=0.005)
    # begin: URCap Program Node
    #   Source: Robotiq_Grippers, 1.8.4.4844, Robotiq Inc.
    #   Type: Gripper
    $ 2348 "Gripper Close (1)"
    if not(gripper_connected[0]):
      popup("Gripper 1 must be connected to run this program.", "No connection", False, True, True)
    end
    if not(rq_is_gripper_activated("1")):
      popup("Gripper 1 is not activated. Go to Installation tab > Gripper to activate it and run the program again.", "Not activated", False, True, True)
    end
    rq_set_pos_spd_for(255, 77, 77, "1")
    rq_wait_pos_spe_for_request(255, 77, 77, "1")
    rq_go_to("1")
    rq_wait("1")
    # end: URCap Program Node
    $ 2349 "CircleMove"
    $ 2350 "ViaPoint_1" "noBreak"

    $ 2351 "Waypoint_57" "breakAfter"
    movec(ViaPoint_1_p, Waypoint_57_p, a=0.3, v=0.05, r=0.005)
    # begin: URCap Program Node
    #   Source: Robotiq_Grippers, 1.8.4.4844, Robotiq Inc.
    #   Type: Gripper
    $ 2352 "Gripper Open (1)"
    if not(gripper_connected[0]):
      popup("Gripper 1 must be connected to run this program.", "No connection", False, True, True)
    end
    if not(rq_is_gripper_activated("1")):
      popup("Gripper 1 is not activated. Go to Installation tab > Gripper to activate it and run the program again.", "Not activated", False, True, True)
    end
    rq_set_pos_spd_for(0, 77, 77, "1")
    rq_wait_pos_spe_for_request(0, 77, 77, "1")
    rq_go_to("1")
    rq_wait("1")
    # end: URCap Program Node
    # begin: URCap Program Node
    #   Source: Robotiq_Grippers, 1.8.4.4844, Robotiq Inc.
    #   Type: Gripper
    $ 2353 "Gripper Open (1)"
    if not(gripper_connected[0]):
      popup("Gripper 1 must be connected to run this program.", "No connection", False, True, True)
    end
    if not(rq_is_gripper_activated("1")):
      popup("Gripper 1 is not activated. Go to Installation tab > Gripper to activate it and run the program again.", "Not activated", False, True, True)
    end
    rq_set_pos_spd_for(0, 77, 77, "1")
    rq_wait_pos_spe_for_request(0, 77, 77, "1")
    rq_go_to("1")
    rq_wait("1")
    # end: URCap Program Node
    $ 2354 "Waypoint_69" "breakAfter"
    movel(Waypoint_69_p, a=1.2, v=0.25, r=0.05)
    $ 2355 "Home (Safe)"
    movej([-1.2302089344500047, -1.2969853503591224, -1.875639182904262, -1.539621866126728, 1.5731943360401213, -2.80099559440227], a=1.3962634015954636, v=1.0471975511965976)
  elif (40 == switch_1):
    $ 2356 "Case 40"
    $ 2396 "Powder dispensing"
    $ 2397 "zero_scale()"
    zero_scale()
    # begin: URCap Program Node
    #   Source: SensoPart VISOR Robotic, 2.0.0, SensoPart Industriesensorik GmbH
    #   Type: VISOR Robotic App
    $ 2398 "VISOR Easy Pick"
    def visorFuncEasyPick_717997():
      # begin: URCap Program Node
      #   Source: SensoPart VISOR Robotic, 2.0.0, SensoPart Industriesensorik GmbH
      #   Type: Easy Pick Setup
      $ 2399 "# 1 Setup" "noBreak"
      local easyPickVisorId = 1
      local easyPickArmMounted = True
      local easyPickSetJob = True
      local easyPickJobName = "Weigh_dispense"
      local easyPickAtImgAcq = False
      local easyPickImgAcqPose = cont_img_pose
      # end: URCap Program Node
      # begin: URCap Program Node
      #   Source: SensoPart VISOR Robotic, 2.0.0, SensoPart Industriesensorik GmbH
      #   Type: Process
      $ 2400 "Process" "noBreak"
      local easyPickObjTaken = False
      local easyPickTrigger = False
      local easyPickPoseIdx = 0
      local easyPickPose = p[0,0,0,0,0,0]
      def easyPickFuncTrigger(visorId, setJob, jobName, arm):
      if (setJob):
        visor_changeJob(visorId, jobName, 6000)
      end
      if (arm):
        visor_trigger(visorId, 6000, "arm")
      else:
        visor_trigger(visorId, 6000)
      end
      global easyPickParts_4=visor_partsFound(visorId)
      visor_easyPickUpdate(visorId, "parts", visor_partsFound(visorId))
      return visor_getPose3d(visorId, 0)
    end
    while (not easyPickObjTaken):
      easyPickTrigger = (easyPickCount_4 >= visor_partsFound(easyPickVisorId)) or (easyPickCount_4 > 9) or (not visor_easyPickCheckIdent("9ccdb7", easyPickVisorId))
      if (easyPickTrigger):
        easyPickCount_4 = 0
      end
      easyPickPoseIdx = easyPickCount_4
      easyPickPose = visor_getPose3d(easyPickVisorId, easyPickPoseIdx)
      visor_easyPickUpdate(easyPickVisorId, "counter", easyPickPoseIdx)
      # begin: URCap Program Node
      #   Source: SensoPart VISOR Robotic, 2.0.0, SensoPart Industriesensorik GmbH
      #   Type: Image Acquisition Pose
      $ 2401 "Image Acquisition Pose" "noBreak"
      if (easyPickTrigger):
        if (not easyPickAtImgAcq):
          movej(pose_trans(easyPickImgAcqPose,p[0.0000,0.0000,-0.0000,0.0000,0.0000,0.0000]),a=1.3963,v=1.0472,t=0.000000,r=0.000000)
          easyPickAtImgAcq = True
        end
        easyPickPose = easyPickFuncTrigger(easyPickVisorId, easyPickSetJob, easyPickJobName, easyPickArmMounted)
      end
      # end: URCap Program Node
      # begin: URCap Program Node
      #   Source: SensoPart VISOR Robotic, 2.0.0, SensoPart Industriesensorik GmbH
      #   Type: Object Detected
      $ 2402 "Object Detected" "noBreak"
      if (visor_partsFound(easyPickVisorId) > 0):
        $ 2403 "Open Gripper" "noBreak"
        $ 2404 "MoveL" "noBreak"
        $ 2405 "Weight_value≔get_weight()" "noBreak"
        global Weight_value=get_weight()
        $ 2406 "Spatula_pick" "noBreak"
        # begin: URCap Program Node
        #   Source: Robotiq_Grippers, 1.8.4.4844, Robotiq Inc.
        #   Type: Gripper
        $ 2407 "Gripper Open (1)" "noBreak"
        if not(gripper_connected[0]):
          popup("Gripper 1 must be connected to run this program.", "No connection", False, True, True)
        end
        if not(rq_is_gripper_activated("1")):
          popup("Gripper 1 is not activated. Go to Installation tab > Gripper to activate it and run the program again.", "Not activated", False, True, True)
        end
        rq_set_pos_spd_for(0, 77, 77, "1")
        rq_wait_pos_spe_for_request(0, 77, 77, "1")
        rq_go_to("1")
        rq_wait("1")
        # end: URCap Program Node
        $ 2408 "Waypoint_53" "noBreak"
        movel(Waypoint_53_p, a=0.6, v=0.15, r=0.05)
        $ 2409 "Spatula_above" "noBreak"
        movel(Spatula_above_p, a=0.6, v=0.15)
        $ 2410 "Spatula_pick" "noBreak"
        movel(Spatula_pick_p, a=0.6, v=0.15)
        # begin: URCap Program Node
        #   Source: Robotiq_Grippers, 1.8.4.4844, Robotiq Inc.
        #   Type: Gripper
        $ 2411 "Gripper Close (1)" "noBreak"
        if not(gripper_connected[0]):
          popup("Gripper 1 must be connected to run this program.", "No connection", False, True, True)
        end
        if not(rq_is_gripper_activated("1")):
          popup("Gripper 1 is not activated. Go to Installation tab > Gripper to activate it and run the program again.", "Not activated", False, True, True)
        end
        rq_set_pos_spd_for(255, 77, 77, "1")
        rq_wait_pos_spe_for_request(255, 77, 77, "1")
        rq_go_to("1")
        rq_wait("1")
        # end: URCap Program Node
        $ 2412 "Spatula_above" "noBreak"
        movel(Spatula_above_p, a=0.6, v=0.15)
        $ 2413 "Popup: Connect the vibration motor" "noBreak"
        popup("Connect the vibration motor", "Message", False, False, blocking=True)
        $ 2414 "tare_scale()" "noBreak"
        tare_scale()
        $ 2415 "PowA_ScoopA" "noBreak"
        movel(PowA_ScoopA_p, a=0.3, v=0.1)
        $ 2416 "scoop" "noBreak"
        global move_thread_flag_2416=0
        thread move_thread_2416():
          enter_critical
          move_thread_flag_2416 = 1
          movel(scoop_p, a=0.6, v=0.15)
          move_thread_flag_2416 = 2
          exit_critical
        end
        move_thread_flag_2416 = 0
        move_thread_han_2416 = run move_thread_2416()
        while (True):
          local targetTcpDirection=get_target_tcp_speed()
          local stepsToRetract=tool_contact(direction=targetTcpDirection)
          if (stepsToRetract > 0):
            kill move_thread_han_2416
            stopl(0.6)
            local backTrackMovement=get_actual_joint_positions_history(stepsToRetract)
            local contactPose=get_forward_kin(backTrackMovement)
            local posDir=[targetTcpDirection[0],targetTcpDirection[1],targetTcpDirection[2]]
            local retractTo=contactPose
            if (norm(posDir) > 1e-6):
              local normalizedPosDir=normalize(posDir)
              local additionalRetraction=p[normalizedPosDir[0] * 0.0, normalizedPosDir[1] * 0.0, normalizedPosDir[2] * 0.0, 0, 0, 0]
              retractTo = pose_sub(contactPose, additionalRetraction)
            end
            movel(retractTo, a=0.6, v=0.1)
            $ 2417 "Until (tool_contact_detection)" "noBreak"
            break
          end
          sleep(1.0E-10)
          if (move_thread_flag_2416 > 1):
            join move_thread_han_2416
            break
          end
          sync()
        end
        $ 2418 "aftr_scoop1" "noBreak"
        movel(aftr_scoop1_p, a=0.5, v=0.2)
        $ 2419 "Set AO[0]=3.0" "noBreak"
        set_standard_analog_out(0, 0.3)
        $ 2420 "Wait: 4.0" "noBreak"
        sleep(4.0)
        $ 2421 "Set AO[0]=0.0" "noBreak"
        set_standard_analog_out(0, 0.0)
        $ 2422 "tilt_angle≔1.5" "noBreak"
        global tilt_angle=1.5
        $ 2423 "ftr_scoop2" "noBreak"
        movel(ftr_scoop2_p, a=0.3, v=0.05)
        $ 2424 "aftr_scoo3" "noBreak"
        movel(aftr_scoo3_p, a=0.3, v=0.075, r=0.01)
        # begin: URCap Program Node
        #   Source: SensoPart VISOR Robotic, 2.0.0, SensoPart Industriesensorik GmbH
        #   Type: Approach Pose
        $ 2425 "Approach Pose" "noBreak"
        movej(pose_trans(easyPickPose,p[0.0000,0.0000,0.0200,0.0000,0.0000,0.0000]),a=0.4363,v=0.3491,t=0.000000,r=0.000000)
        # end: URCap Program Node
        # begin: URCap Program Node
        #   Source: SensoPart VISOR Robotic, 2.0.0, SensoPart Industriesensorik GmbH
        #   Type: Target Pose
        $ 2426 "Target Pose" "noBreak"
        movel(pose_trans(easyPickPose,p[0.0000,0.0000,-0.0000,0.0000,0.0000,0.0000]),a=0.1000,v=0.0500,t=0.000000,r=0.000000)
        # end: URCap Program Node
        $ 2427 "Close Gripper" "noBreak"
        $ 2428 "dispense_pos≔get_actual_tcp_pose()" "noBreak"
        global dispense_pos= get_actual_tcp_pose ()
        $ 2429 "MoveL" "noBreak"
        $ 2430 "Start_thread≔ True " "noBreak"
        global Start_thread=  True
        $ 2431 "vib_mot_thread≔ True " "noBreak"
        global vib_mot_thread=  True
        $ 2432 "Wait: 0.5" "noBreak"
        sleep(0.5)
        $ 2433 "Loop Weight_value≤Target_weight and tilt_angle≥1.1" "noBreak"
        thread Thread_while_2433():
          while (True):
            $ 2434 "current_error≔Target_weight-Weight_value" "noBreak"
            global current_error=Target_weight-Weight_value
            $ 2435 "Integral_error≔Integral_error+current_error*dt" "noBreak"
            global Integral_error=Integral_error+current_error*dt
            $ 2436 "derivative≔(current_error-previous_error)/dt" "noBreak"
            global derivative=(current_error-previous_error)/dt
            $ 2437 "tilt_increment≔(kp*current_error)+(ki*Integral_error)+(kd*derivative)" "noBreak"
            global tilt_increment=(kp*current_error)+(ki*Integral_error)+(kd*derivative)
            $ 2438 "current_pose≔get_actual_tcp_pose()" "noBreak"
            global current_pose= get_actual_tcp_pose ()
            $ 2439 "tilt_angle≔current_pose[4]" "noBreak"
            global tilt_angle=current_pose[4]
            $ 2440 "If tilt_increment>0.1" "noBreak"
            global thread_flag_2440=0
            thread Thread_if_2440():
              $ 2441 "tilt_increment≔0.05" "noBreak"
              global tilt_increment=0.05
              thread_flag_2440 = 1
            end
            if (tilt_increment>0.1):
              global thread_handler_2440=run Thread_if_2440()
              while (thread_flag_2440 == 0):
                if not(tilt_increment>0.1):
                  kill thread_handler_2440
                  thread_flag_2440 = 2
                else:
                  sync()
                end
              end
            else:
              thread_flag_2440 = 2
            end
            $ 2442 "tilt_pose≔pose_trans(current_pose, p[(-tilt_increment/5), 0, 0, 0, -tilt_increment, 0])" "noBreak"
            global tilt_pose=pose_trans(current_pose, p[(-tilt_increment/5), 0, 0, 0, -tilt_increment, 0])
            $ 2443 "movel(tilt_pose, a=0.025, v=0.015, r=0.00001)" "noBreak"
            movel(tilt_pose, a=0.025, v=0.015, r=0.00001)
            $ 2444 "previous_error≔current_error" "noBreak"
            global previous_error=current_error
          end
        end
        if (Weight_value <= Target_weight  and  tilt_angle >= 1.1):
          global thread_handler_2433=run Thread_while_2433()
          while (Weight_value <= Target_weight  and  tilt_angle >= 1.1):
            sync()
          end
          kill thread_handler_2433
        end
        $ 2445 "Start_thread≔ False " "noBreak"
        global Start_thread=  False
        $ 2447 "Weight_value≔get_weight()" "noBreak"
        global Weight_value=get_weight()
        $ 2448 "Wait: 0.5" "noBreak"
        sleep(0.5)
        $ 2449 "vib_mot_thread≔ False " "noBreak"
        global vib_mot_thread=  False
        $ 2450 "MoveL" "noBreak"
        $ 2451 "dispense_pos" "noBreak"
        movel(dispense_pos, a=0.2, v=0.05)
        $ 2452 "Integral_error≔0" "noBreak"
        global Integral_error=0
        $ 2453 "current_error≔0" "noBreak"
        global current_error=0
        $ 2454 "previous_error≔0" "noBreak"
        global previous_error=0
        $ 2455 "Set AO[0]=0.0" "noBreak"
        set_standard_analog_out(0, 0.0)
        # begin: URCap Program Node
        #   Source: SensoPart VISOR Robotic, 2.0.0, SensoPart Industriesensorik GmbH
        #   Type: Exit Pose
        $ 2456 "Exit Pose" "noBreak"
        movel(pose_trans(easyPickPose,p[0.0000,0.0000,-0.0000,0.0000,0.0000,0.0000]),a=0.5000,v=0.2500,t=0.000000,r=0.000000)
        # end: URCap Program Node
        easyPickObjTaken = True
      end
      # end: URCap Program Node
      # begin: URCap Program Node
      #   Source: SensoPart VISOR Robotic, 2.0.0, SensoPart Industriesensorik GmbH
      #   Type: No Object Detected
      $ 2457 "No Object Detected" "noBreak"
      if (visor_partsFound(easyPickVisorId) < 1):
        $ 2458 "Popup: No weigh scale detected" "noBreak"
        popup("No weigh scale detected", "Message", False, False, blocking=True)
        else:
      end
      # end: URCap Program Node
    end
    easyPickCount_4 = easyPickCount_4 + 1
    visor_easyPickUpdate(easyPickVisorId, "counter", easyPickCount_4)
    visor_easyPickSetIdent("9ccdb7", easyPickVisorId)
    # end: URCap Program Node
  end
  visorFuncEasyPick_717997()
  # end: URCap Program Node
  $ 2459 "powder dispensing"
  $ 2461 "Loop Weight_value<Target_weight"
  while (Weight_value<Target_weight):
    $ 2462 "MoveL"
    $ 2463 "Waypoint_75" "breakAfter"
    movel(Waypoint_75_p, a=0.3, v=0.05, r=0.05)
    $ 2464 "Waypoint_71" "breakAfter"
    movel(Waypoint_71_p, a=0.3, v=0.05)
    $ 2465 "Waypoint_83" "breakAfter"
    movel(Waypoint_83_p, a=0.3, v=0.05)
    $ 2466 "Waypoint_73" "breakAfter"
    movel(Waypoint_73_p, a=0.3, v=0.05, r=0.005)
    $ 2467 "scoop" "breakAfter"
    global move_thread_flag_2467=0
    thread move_thread_2467():
      enter_critical
      move_thread_flag_2467 = 1
      movel(scoop_p, a=0.3, v=0.1)
      move_thread_flag_2467 = 2
      exit_critical
    end
    move_thread_flag_2467 = 0
    move_thread_han_2467 = run move_thread_2467()
    while (True):
      local targetTcpDirection=get_target_tcp_speed()
      local stepsToRetract=tool_contact(direction=targetTcpDirection)
      if (stepsToRetract > 0):
        kill move_thread_han_2467
        stopl(3.0)
        local backTrackMovement=get_actual_joint_positions_history(stepsToRetract)
        local contactPose=get_forward_kin(backTrackMovement)
        local posDir=[targetTcpDirection[0],targetTcpDirection[1],targetTcpDirection[2]]
        local retractTo=contactPose
        if (norm(posDir) > 1e-6):
          local normalizedPosDir=normalize(posDir)
          local additionalRetraction=p[normalizedPosDir[0] * 0.0, normalizedPosDir[1] * 0.0, normalizedPosDir[2] * 0.0, 0, 0, 0]
          retractTo = pose_sub(contactPose, additionalRetraction)
        end
        movel(retractTo, a=3.0, v=0.1)
        $ 2468 "Until (tool_contact_detection)"
        break
      end
      sleep(1.0E-10)
      if (move_thread_flag_2467 > 1):
        join move_thread_han_2467
        break
      end
      sync()
    end
    $ 2469 "aftr_scoop1" "breakAfter"
    movel(aftr_scoop1_p, a=0.3, v=0.05)
    $ 2470 "Set AO[0]=3.0"
    set_standard_analog_out(0, 0.3)
    $ 2471 "Wait: 3.0"
    sleep(3.0)
    $ 2472 "Set AO[0]=0.0"
    set_standard_analog_out(0, 0.0)
    $ 2473 "ftr_scoop2" "breakAfter"
    movel(ftr_scoop2_p, a=0.3, v=0.05)
    $ 2474 "aftr_scoo3" "breakAfter"
    movel(aftr_scoo3_p, a=0.3, v=0.05)
    $ 2475 "MoveL"
    $ 2476 "Start_thread≔ True "
    global Start_thread=  True
    $ 2477 "dispense_pos" "breakAfter"
    movel(dispense_pos, a=0.2, v=0.05)
    $ 2478 "tilt_angle≔1.5"
    global tilt_angle=1.5
    $ 2479 "vib_mot_thread≔ True "
    global vib_mot_thread=  True
    $ 2480 "Wait: 0.5"
    sleep(0.5)
    $ 2481 "Loop Weight_value≤Target_weight and tilt_angle≥1.1"
    thread Thread_while_2481():
      while (True):
        $ 2482 "current_error≔Target_weight-Weight_value"
        global current_error=Target_weight-Weight_value
        $ 2483 "Integral_error≔Integral_error+current_error*dt"
        global Integral_error=Integral_error+current_error*dt
        $ 2484 "derivative≔(current_error-previous_error)/dt"
        global derivative=(current_error-previous_error)/dt
        $ 2485 "tilt_increment≔(kp*current_error)+(ki*Integral_error)+(kd*derivative)"
        global tilt_increment=(kp*current_error)+(ki*Integral_error)+(kd*derivative)
        $ 2486 "current_pose≔get_actual_tcp_pose()"
        global current_pose= get_actual_tcp_pose ()
        $ 2487 "tilt_angle≔current_pose[4]"
        global tilt_angle=current_pose[4]
        $ 2488 "If tilt_increment>0.1"
        global thread_flag_2488=0
        thread Thread_if_2488():
          $ 2489 "tilt_increment≔0.05"
          global tilt_increment=0.05
          thread_flag_2488 = 1
        end
        if (tilt_increment>0.1):
          global thread_handler_2488=run Thread_if_2488()
          while (thread_flag_2488 == 0):
            if not(tilt_increment>0.1):
              kill thread_handler_2488
              thread_flag_2488 = 2
            else:
              sync()
            end
          end
        else:
          thread_flag_2488 = 2
        end
        $ 2490 "tilt_pose≔pose_trans(current_pose, p[(-tilt_increment/5), 0, 0, 0, -tilt_increment, 0])"
        global tilt_pose=pose_trans(current_pose, p[(-tilt_increment/5), 0, 0, 0, -tilt_increment, 0])
        $ 2491 "movel(tilt_pose, a=0.020, v=0.010, r=0.00001)"
        movel(tilt_pose, a=0.020, v=0.010, r=0.00001)
        $ 2492 "previous_error≔current_error"
        global previous_error=current_error
        $ 2493 "Wait: 0.01"
        sleep(0.01)
      end
    end
    if (Weight_value <= Target_weight  and  tilt_angle >= 1.1):
      global thread_handler_2481=run Thread_while_2481()
      while (Weight_value <= Target_weight  and  tilt_angle >= 1.1):
        sync()
      end
      kill thread_handler_2481
    end
    $ 2494 "Start_thread≔ False "
    global Start_thread=  False
    $ 2495 "vib_mot_thread≔ False "
    global vib_mot_thread=  False
    $ 2497 "Weight_value≔get_weight()"
    global Weight_value=get_weight()
    $ 2498 "Set AO[0]=0.0"
    set_standard_analog_out(0, 0.0)
    $ 2500 "Wait: 0.5"
    sleep(0.5)
    $ 2501 "MoveL"
    $ 2502 "dispense_pos" "breakAfter"
    movel(dispense_pos, a=0.1, v=0.05)
    $ 2503 "Integral_error≔0"
    global Integral_error=0
    $ 2504 "current_error≔0"
    global current_error=0
    $ 2505 "previous_error≔0"
    global previous_error=0
  end
  $ 2506 "MoveL"
  $ 2507 "aftr_scoo3" "breakAfter"
  movel(aftr_scoo3_p, a=0.3, v=0.1)
  $ 2508 "ftr_scoop2" "breakAfter"
  movel(ftr_scoop2_p, a=0.4, v=0.1)
  $ 2509 "aftr_scoop1" "breakAfter"
  movel(aftr_scoop1_p, a=0.4, v=0.1)
  $ 2510 "aftr_disp4" "breakAfter"
  movel(aftr_disp4_p, a=0.3, v=0.05)
  $ 2511 "Set AO[0]=3.0"
  set_standard_analog_out(0, 0.3)
  $ 2512 "Wait: 2.0"
  sleep(2.0)
  $ 2513 "Set AO[0]=0.0"
  set_standard_analog_out(0, 0.0)
  $ 2514 "Waypoint_84" "breakAfter"
  movel(Waypoint_84_p, a=0.3, v=0.075, r=0.005)
  $ 2515 "Waypoint_54" "breakAfter"
  movel(Waypoint_54_p, a=0.3, v=0.075, r=0.05)
  $ 2516 "Spatula_above" "breakAfter"
  movel(Spatula_above_p, a=0.3, v=0.1, r=0.003)
  $ 2517 "Waypoint_58" "breakAfter"
  movel(Waypoint_58_p, a=1.2, v=0.25)
  $ 2518 "Waypoint_59" "breakAfter"
  movel(Waypoint_59_p, a=0.3, v=0.1)
  $ 2519 "Popup: Disconnect the vibration motor"
  popup("Disconnect the vibration motor", "Message", False, False, blocking=True)
  $ 2520 "Waypoint_72" "breakAfter"
  movel(Waypoint_72_p, a=0.3, v=0.1)
  # begin: URCap Program Node
  #   Source: Robotiq_Grippers, 1.8.4.4844, Robotiq Inc.
  #   Type: Gripper
  $ 2521 "Gripper Open (1)"
  if not(gripper_connected[0]):
    popup("Gripper 1 must be connected to run this program.", "No connection", False, True, True)
  end
  if not(rq_is_gripper_activated("1")):
    popup("Gripper 1 is not activated. Go to Installation tab > Gripper to activate it and run the program again.", "Not activated", False, True, True)
  end
  rq_set_pos_spd_for(0, 77, 77, "1")
  rq_wait_pos_spe_for_request(0, 77, 77, "1")
  rq_go_to("1")
  rq_wait("1")
  # end: URCap Program Node
  $ 2522 "Spatula_above" "breakAfter"
  movel(Spatula_above_p, a=1.2, v=0.25)
  $ 2524 "Cap the container"
  $ 2525 "MoveL"
  $ 2526 "Waypoint_69" "breakAfter"
  movel(Waypoint_69_p, a=1.2, v=0.25, r=0.05)
  $ 2527 "Waypoint_57" "breakAfter"
  movel(Waypoint_57_p, a=0.6, v=0.15)
  # begin: URCap Program Node
  #   Source: Robotiq_Grippers, 1.8.4.4844, Robotiq Inc.
  #   Type: Gripper
  $ 2528 "Gripper Close (1)"
  if not(gripper_connected[0]):
    popup("Gripper 1 must be connected to run this program.", "No connection", False, True, True)
  end
  if not(rq_is_gripper_activated("1")):
    popup("Gripper 1 is not activated. Go to Installation tab > Gripper to activate it and run the program again.", "Not activated", False, True, True)
  end
  rq_set_pos_spd_for(255, 77, 77, "1")
  rq_wait_pos_spe_for_request(255, 77, 77, "1")
  rq_go_to("1")
  rq_wait("1")
  # end: URCap Program Node
  $ 2529 "Waypoint_68" "breakAfter"
  movel(Waypoint_68_p, a=0.6, v=0.15, r=0.005)
  $ 2530 "Waypoint_67" "breakAfter"
  movel(Waypoint_67_p, a=0.6, v=0.15, r=0.005)
  $ 2531 "Waypoint_66" "breakAfter"
  movel(Waypoint_66_p, a=0.6, v=0.15, r=0.005)
  $ 2532 "Waypoint_52" "breakAfter"
  movel(Waypoint_52_p, a=1.2, v=0.25)
  # begin: URCap Program Node
  #   Source: Robotiq_Grippers, 1.8.4.4844, Robotiq Inc.
  #   Type: Gripper
  $ 2533 "Gripper Open (1)"
  if not(gripper_connected[0]):
    popup("Gripper 1 must be connected to run this program.", "No connection", False, True, True)
  end
  if not(rq_is_gripper_activated("1")):
    popup("Gripper 1 is not activated. Go to Installation tab > Gripper to activate it and run the program again.", "Not activated", False, True, True)
  end
  rq_set_pos_spd_for(0, 77, 77, "1")
  rq_wait_pos_spe_for_request(0, 77, 77, "1")
  rq_go_to("1")
  rq_wait("1")
  # end: URCap Program Node
  $ 2534 "Tilt_above" "breakAfter"
  movel(Tilt_above_p, a=1.2, v=0.25)
  $ 2535 "Tilt_place" "breakAfter"
  movel(Tilt_place_p, a=0.3, v=0.05)
  # begin: URCap Program Node
  #   Source: Robotiq_Grippers, 1.8.4.4844, Robotiq Inc.
  #   Type: Gripper
  $ 2536 "Gripper Close (1)"
  if not(gripper_connected[0]):
    popup("Gripper 1 must be connected to run this program.", "No connection", False, True, True)
  end
  if not(rq_is_gripper_activated("1")):
    popup("Gripper 1 is not activated. Go to Installation tab > Gripper to activate it and run the program again.", "Not activated", False, True, True)
  end
  rq_set_pos_spd_for(255, 77, 77, "1")
  rq_wait_pos_spe_for_request(255, 77, 77, "1")
  rq_go_to("1")
  rq_wait("1")
  # end: URCap Program Node
  $ 2537 "Tilt_above" "breakAfter"
  movel(Tilt_above_p, a=0.3, v=0.1)
  $ 2538 "OP_PowderA_abov" "breakAfter"
  movel(OP_PowderA_abov_p, a=0.3, v=0.05)
  $ 2539 "Set GRP_3F_Open=On"
  set_standard_digital_out(5, True)
  $ 2540 "Wait: 0.5"
  sleep(0.5)
  $ 2541 "OP_PowderA_pick" "breakAfter"
  movel(OP_PowderA_pick_p, a=0.3, v=0.1)
  $ 2542 "Set GRP_3F_Open=Off"
  set_standard_digital_out(5, False)
  $ 2543 "Wait: 0.5"
  sleep(0.5)
  # begin: URCap Program Node
  #   Source: Robotiq_Grippers, 1.8.4.4844, Robotiq Inc.
  #   Type: Gripper
  $ 2544 "Gripper Open (1)"
  if not(gripper_connected[0]):
    popup("Gripper 1 must be connected to run this program.", "No connection", False, True, True)
  end
  if not(rq_is_gripper_activated("1")):
    popup("Gripper 1 is not activated. Go to Installation tab > Gripper to activate it and run the program again.", "Not activated", False, True, True)
  end
  rq_set_pos_spd_for(0, 77, 77, "1")
  rq_wait_pos_spe_for_request(0, 77, 77, "1")
  rq_go_to("1")
  rq_wait("1")
  # end: URCap Program Node
  $ 2545 "OP_PowderA_abov" "breakAfter"
  movel(OP_PowderA_abov_p, a=1.2, v=0.25)
  $ 2546 "OP_PowderA2" "breakAfter"
  movel(OP_PowderA2_p, a=1.2, v=0.25)
  $ 2547 "Home (Safe)"
  movej([-1.2302089344500047, -1.2969853503591224, -1.875639182904262, -1.539621866126728, 1.5731943360401213, -2.80099559440227], a=1.3962634015954636, v=1.0471975511965976)
  $ 2548 "Cap_above" "breakAfter"
  movel(Cap_above_p, a=1.2, v=0.25)
  # begin: URCap Program Node
  #   Source: Robotiq_Grippers, 1.8.4.4844, Robotiq Inc.
  #   Type: Gripper
  $ 2549 "Gripper Open (1)"
  if not(gripper_connected[0]):
    popup("Gripper 1 must be connected to run this program.", "No connection", False, True, True)
  end
  if not(rq_is_gripper_activated("1")):
    popup("Gripper 1 is not activated. Go to Installation tab > Gripper to activate it and run the program again.", "Not activated", False, True, True)
  end
  rq_set_pos_spd_for(0, 77, 77, "1")
  rq_wait_pos_spe_for_request(0, 77, 77, "1")
  rq_go_to("1")
  rq_wait("1")
  # end: URCap Program Node
  $ 2550 "Cap_Place" "breakAfter"
  movel(Cap_Place_p, a=1.2, v=0.25)
  # begin: URCap Program Node
  #   Source: Robotiq_Grippers, 1.8.4.4844, Robotiq Inc.
  #   Type: Gripper
  $ 2551 "Gripper Move22mm (1)"
  if not(gripper_connected[0]):
    popup("Gripper 1 must be connected to run this program.", "No connection", False, True, True)
  end
  if not(rq_is_gripper_activated("1")):
    popup("Gripper 1 is not activated. Go to Installation tab > Gripper to activate it and run the program again.", "Not activated", False, True, True)
  end
  rq_set_pos_spd_for(145, 77, 77, "1")
  rq_wait_pos_spe_for_request(145, 77, 77, "1")
  rq_go_to("1")
  rq_wait("1")
  # end: URCap Program Node
  $ 2552 "Cap_above" "breakAfter"
  movel(Cap_above_p, a=1.2, v=0.25, r=0.05)
  $ 2553 "Waypoint_82" "breakAfter"
  movel(Waypoint_82_p, a=1.2, v=0.25)
  $ 2554 "Waypoint_81" "breakAfter"
  movel(Waypoint_81_p, a=0.3, v=0.1)
  $ 2556 "Cap"
  $ 2557 "Action_Info≔'capping'"
  global Action_Info="capping"
  $ 2558 "Set GRP_3F_Enable=On"
  set_standard_digital_out(4, True)
  $ 2559 "Set GRP_3F_Cap=On"
  set_standard_digital_out(2, True)
  $ 2562 "Waypoint_77" "breakAfter"
  movel(Waypoint_77_p, t=4.0)
  $ 2563 "Set GRP_3F_Cap=Off"
  set_standard_digital_out(2, False)
  $ 2564 "Set GRP_3F_Enable=Off"
  set_standard_digital_out(4, False)
  # begin: URCap Program Node
  #   Source: Robotiq_Grippers, 1.8.4.4844, Robotiq Inc.
  #   Type: Gripper
  $ 2565 "Gripper Open (1)"
  if not(gripper_connected[0]):
    popup("Gripper 1 must be connected to run this program.", "No connection", False, True, True)
  end
  if not(rq_is_gripper_activated("1")):
    popup("Gripper 1 is not activated. Go to Installation tab > Gripper to activate it and run the program again.", "Not activated", False, True, True)
  end
  rq_set_pos_spd_for(0, 77, 77, "1")
  rq_wait_pos_spe_for_request(0, 77, 77, "1")
  rq_go_to("1")
  rq_wait("1")
  # end: URCap Program Node
  $ 2566 "Waypoint_82" "breakAfter"
  movel(Waypoint_82_p, a=1.2, v=0.25)
  $ 2567 "Home (Safe)"
  movej([-1.2302089344500047, -1.2969853503591224, -1.875639182904262, -1.539621866126728, 1.5731943360401213, -2.80099559440227], a=1.3962634015954636, v=1.0471975511965976)
  end
  $ 2568 "'=========='"
  # '=========='
  $ 2569 "PostSettings"
  $ 2570 "'ADD ADDITIONAL CHECKS'"
  # 'ADD ADDITIONAL CHECKS'
  end
  $ 2 "BeforeStart"
  $ 3 "Scripts"
  $ 4 "Script: 001 SCRIPT Errors and Warnings Deifnes V0.2.script"

  #*****************************************************
  # customer          :   UK Essen
  # project name      :   P1132
  #****************************************************
  # controller        :
  # software          :
  #****************************************************
  # author            :   E.Petrichenko
  # Copyright (c)     :   United Robotics Group Health and Food GmbH
  #                       An der Riede 2
  #                       28816 Stuhr
  #                       Germany
  #****************************************************
  # description       :   centrifuge actions for the application
  # version:      	:   0.1
  # created           :   22.08.2024
  # updated           :
  #****************************************************
  # modifications     :
  #
  # date              :
  # name              :
  # reason            :
  #****************************************************


  #################################### VARIABLES DEFINITIONS ###################################

  ERROR_POSE_NOT_REACHABLE = 1002
  ERROR_ROBOT_ARM_NOT_IN_HOME_POSE = 1006
  ERROR_NO_OBJECT_TO_PICK = 1010
  ERROR_NOT_DOCKED = 2003
  ERROR_NOT_REACHABLE_TARGET = 2007
  ERROR_CHARGING_NOT_STARTED = 2008
  ERROR_AMR_WRONG_MODE = 2009
  ERROR_UNKNOWN_POSE = 2010
  ERROR_NO_LANDMARK = 3002
  ERROR_WRONG_ORDER = 4002
  ERROR_CENTRIFUGE_CONNECTION = 5001
  ERROR_CENTRIFUGE_POWER = 5002
  ERROR_CENTRIFUGE = 5003
  ERROR_CENTRIFUGE_LID = 5004
  ERROR_CANNOT_OPEN_HATCH = 5006
  ERROR_CANNOT_CLOSE_HATCH = 5008
  ERROR_CANNOT_ROTATE = 5010
  ERROR_CANNOT_START = 5011
  ERROR_WRONG_KEY_POSE = 5012
  ERROR_MISSIING_CENTRACK = 5013

  WARNING_POSE_NOT_REACHABLE = 1002
  WARNING_BATTERY_LEVEL = 2002
  WARNING_NOT_REACHABLE_TARGET = 2007


  ERROR = struct(
      FLAG = False,
      ID = 0,
      MSG = "")

  WARNING = struct(
      FLAG = False,
      ID = 0,
      MSG = "")


  #################################### FUNCTIONS ###################################

  def set_error(error_id):
      ERROR.ID = error_id
      if (ERROR.ID == 0):
          ERROR.FLAG = False
          ERROR.MSG = ""
      else:
          ERROR.FLAG = True
          if(ERROR.ID == ERROR_POSE_NOT_REACHABLE):
              ERROR.MSG = "Pose is not reachable"
          elif(ERROR.ID == ERROR_NO_OBJECT_TO_PICK):
              ERROR.MSG = "No object to pick"
          elif(ERROR.ID == ERROR_NO_LANDMARK):
              ERROR.MSG = "No landmark detected"
          elif(ERROR.ID == ERROR_ROBOT_ARM_NOT_IN_HOME_POSE):
              ERROR.MSG = "Robot arm cannot go to home pose"
          elif(ERROR.ID == ERROR_AMR_WRONG_MODE):
              ERROR.MSG = "AMR is in the wrong mode"
          elif(ERROR.ID == ERROR_NOT_DOCKED):
              ERROR.MSG = "Could not dock to the charger"
          elif(ERROR.ID == ERROR_NOT_REACHABLE_TARGET):
              ERROR.MSG = "Could not reach the target"
          elif(ERROR.ID == ERROR_CHARGING_NOT_STARTED):
              ERROR.MSG = "Could not start charging"
          elif(ERROR.ID == ERROR_UNKNOWN_POSE):
              ERROR.MSG = "Unknown navigation target"
          elif(ERROR.ID == ERROR_CANNOT_OPEN_HATCH):
              ERROR.MSG = "Centrifuge Cannot open the hatch"
          elif(ERROR.ID == ERROR_CENTRIFUGE_CONNECTION):
              ERROR.MSG = "Cannot reach centrifuge"
          elif (ERROR.ID == ERROR_CANNOT_CLOSE_HATCH):
              ERROR.MSG = "Centrifuge Cannot close the hatch"
          elif (ERROR.ID == ERROR_CANNOT_START):
              ERROR.MSG = "Centrifuge Cannot start"
          elif (ERROR.ID == ERROR_CANNOT_ROTATE):
              ERROR.MSG = "Centrifuge Cannot rotate the rotor"
          elif (ERROR.ID == ERROR_WRONG_ORDER):
              ERROR.MSG = "Wrong parameter was recieved"
          elif (ERROR.ID == ERROR_CENTRIFUGE):
              ERROR.MSG = "Centrifuge is in Error"
          elif (ERROR.ID == ERROR_WRONG_KEY_POSE):
              ERROR.MSG = "Key is in the wrong position"
          elif(ERROR.ID == ERROR_MISSIING_CENTRACK):
              ERROR.MSG = "Missing rack for centrifuge set"
          elif(ERROR.ID == ERROR_CENTRIFUGE_POWER):
              ERROR.MSG = "Centrifuge is turned off"
          elif(ERROR.ID == ERROR_CENTRIFUGE_LID):
              ERROR.MSG = "Lid of the centrifuge is opened"
          else:
              ERROR.MSG = "Unknown code"
          end
          textmsg("ERROR:",ERROR)
      end
  end

  def set_warning(warning_id):
      WARNING.ID = warning_id
      if (WARNING.ID == 0):
          WARNING.FLAG = False
          WARNING.MSG = ""
      else:
          WARNING.FLAG = True
          if(WARNING.ID == WARNING_POSE_NOT_REACHABLE):
              WARNING.MSG = "Pose is not reachable"
          elif(WARNING.ID == WARNING_BATTERY_LEVEL):
              WARNING.MSG = "Batery level dropped to a certain level"
          elif(WARNING.ID == WARNING_NOT_REACHABLE_TARGET):
              WARNING.MSG = "Not reachable location of AMR"
          else:
              WARNING.MSG = "Unknown code"
          end
          textmsg("WARNING:",WARNING)
      end
  end


  def reset_error():
    ERROR.ID = 0
    ERROR.FLAG = False
    ERROR.MSG = ""
  end


  def reset_warning():
      WARNING.ID = 0
      WARNING.FLAG = False
      WARNING.MSG = ""
    end
  $ 5 "Script: SCRIPT uGO V7.11.1.script"
  #*****************************************************
  # customer          :
  # project name      :   Standard Application
  #****************************************************
  # controller        :
  # software          :
  #****************************************************
  # author            :   P. Koehnke
  # Copyright (c)     :   United Robotics Group
  #                       An der Riede 2
  #                       28816 Stuhr
  #                       Germany
  #****************************************************
  # description       :   interface for uGo
  # version:      	:   6.0
  # created           :   21.04.2022
  # updated           :
  #****************************************************
  # modifications     :   add new rpc-functions to interchange more data
  #
  # date              :   2024-02-29
  # name              :   P. Koehnke
  # reason            :   implemtentation of PackML behavoiur in uGO
  #****************************************************
  #****************************************************
  # modifications     :   add reflecting the UID of the uGO task back to uGO
  #
  # date              :   2024-07-02
  # name              :   P. Koehnke
  # reason            :   be sure to finish the right tasks
  #****************************************************

  # available rpc-functions:
  #.on('con_check', (err, _params, callback) => callback(err, this.con_check()))
  #.on('read_input', (err, params, callback) => callback(err, this.read_input(params[0], params[1])))
  #.on('write_output', (err, params, callback) => callback(err, this.write_output(params[0], params[1], params[2])))
  #.on('read_status', (err, params, callback) => callback(err, this.read_status(params[0])))
  #.on('write_status', (err, params, callback) => callback(err, this.write_status(params[0], params[1])))
  #.on('send_template', (err, params, callback) => callback(err, this.receive_state(params[0])))
  #.on('receive_event', (err, params, callback) => callback(err, this.send_event()))
  #.on('send_state', (err, params, callback) => callback(err, this.receive_state(params[0])))
  #.on('send_error', (err, params, callback) => callback(err, this.receive_error(params[0])))
  #.on('NotFound', (methodCalled, params) => LOG.warn('Method "', methodCalled, '" does not exist. ', { params }));

  # =======================================================================
  local IDX_CMD_STOP = 0
  local IDX_CMD_RESET = 1
  local IDX_CMD_START = 2
  local IDX_CMD_HOLD = 3
  local IDX_CMD_UNHOLD = 4
  local IDX_CMD_SUSPEND = 5
  local IDX_CMD_UNSUSPEND = 6
  local IDX_CMD_ABORT = 7
  local IDX_CMD_CLEAR = 8
  local IDX_FNC_FREEDRIVE = 9

  # uGo specific declarations
  global UGO_Request_ID = ""
  global UGO_UNIT_Task = ""
  global UGO_Task_ID = 0
  global UGO_Event = ""
  local UGO_Enable_Control = False
  local UGO = rpc_factory("xmlrpc", "http://192.168.12.120:8080")
  local UGO_Ctrl_Cmd = [False, False, False, False, False, False, False, False, False, False]

  local UGO_AMR_Pos = struct(position_identifier=0, x1=0, x2=0, y1=0, y2=0, theta1=0, theta2=0)
  local UGO_EOAT = struct(object_picked=False)

  def ugo_init(enable=True, rpc_address="http://192.168.12.120:8080"):
      # connection with uGo
      if enable:
          UGO = rpc_factory("xmlrpc", rpc_address)
          UGO_Enable_Control = True
      else:
          UGO_Enable_Control = False
      end
  end

  def ugo_event_controller():
      # interpret the given command and map it to the internal commands
      if UGO_Enable_Control:
          UGO_Event = UGO.receive_event()
      end

      UGO_Ctrl_Cmd[IDX_CMD_STOP] = (UGO_Event == "stop")
      UGO_Ctrl_Cmd[IDX_CMD_RESET] = (UGO_Event == "reset")
      UGO_Ctrl_Cmd[IDX_CMD_START] = (UGO_Event == "start")
      UGO_Ctrl_Cmd[IDX_CMD_HOLD] = (UGO_Event == "hold")
      UGO_Ctrl_Cmd[IDX_CMD_UNHOLD] = (UGO_Event == "un_hold")
      UGO_Ctrl_Cmd[IDX_CMD_SUSPEND] = (UGO_Event == "suspend")
      UGO_Ctrl_Cmd[IDX_CMD_UNSUSPEND] = (UGO_Event == "un_suspend")
      UGO_Ctrl_Cmd[IDX_CMD_ABORT] = (UGO_Event == "abort")
      UGO_Ctrl_Cmd[IDX_CMD_CLEAR] = (UGO_Event == "clear")
      UGO_Ctrl_Cmd[IDX_FNC_FREEDRIVE] = (UGO_Event == "freedrive")

      return UGO_Ctrl_Cmd
  end

  def ugo_translate_pml_state():
      # translate the current PML State to a string
      if (STATE == 1):
          return "STOPPING"
      elif (STATE == 2):
          return "STOPPED"
      elif (STATE == 3):
          return "RESETTING"
      elif (STATE == 4):
          return "IDLE"
      elif (STATE == 5):
          return "STARTING"
      elif (STATE == 6):
          return "EXECUTE"
      elif (STATE == 7):
          return "COMPLETING"
      elif (STATE == 8):
          return "COMPLETE"
      elif (STATE == 9):
          return "HOLDING"
      elif (STATE == 10):
          return "HELD"
      elif (STATE == 11):
          return "UNHOLDING"
      elif (STATE == 12):
          return "SUSPENDING"
      elif (STATE == 13):
          return "SUSPENDED"
      elif (STATE == 14):
          return "UNSUSPENDING"
      elif (STATE == 15):
          return "ABORTING"
      elif (STATE == 16):
          return "ABORTED"
      elif (STATE == 17):
          return "CLEARING"
      else:
          return "UNKNOWN"
      end
  end

  def ugo_update_outputs():
      #Update the outputs to uGo via xmplrpc service
      UGO.write_status("ROB_Skill", UGO_UNIT_Task)
      UGO.write_status("ROB_Battery", AMR_Battery)
      UGO.write_status("ROB_Gripper", OBJ_Picked)
      UGO.send_state(ugo_translate_pml_state(), UGO_UNIT_Task)
      UGO.send_error(ERROR.ID)
      #UGO.send_position(AMR_Position)
  end

  def ugo_get_task():
      # get the actual task to work on
      # added: reflecting the UID of the task back to uGO
      UGO_UNIT_Task = UGO.read_status("DSH_Workflow")
      if (UGO_UNIT_Task != ""):
          UGO_Request_ID = str_sub(UGO_UNIT_Task, 0, 39)
          UGO_Task_ID = to_num(str_sub(UGO_UNIT_Task, 40, 2))
          #ugo_tasks()
          return UGO_Task_ID
      else:
          return 0
      end
  end

  def ugo_pml_stopping():
      return True
  end

  def ugo_pml_resetting():
      ugo_get_task()
      if (UGO_UNIT_Task == ""):
          UGO_Request_ID = ""
          UGO_Task_ID = 0
          return True
      end
      return False
  end

  def ugo_pml_starting():
      #UGO_Task_Content = UGO.receive_task()
      return (UGO_UNIT_Task != "")
  end

  def ugo_pml_holding():
      return True
  end

  def ugo_pml_unholding():
      return True
  end

  def ugo_pml_suspending():
      return True
  end

  def ugo_pml_unsuspending():
      return True
  end

  def ugo_pml_completing():
      return True
  end

  def ugo_pml_aborting():
      return True
  end

  def ugo_pml_clearing():
      return True
  end

  # =======================================================================
  # end of uGO script
  # =======================================================================
  $ 7 "Script: SCRIPT PackML V1.2.1.script"
  # PackML

  IO_ADDRESS_CMD_STOP = 1
  IO_ADDRESS_CMD_RESET = 7
  IO_ADDRESS_CMD_START = 0

  EXT_ADDRESS_CMD_STOP = 0
  EXT_ADDRESS_CMD_RESET = 1
  EXT_ADDRESS_CMD_START = 2
  EXT_ADDRESS_CMD_HOLD = 3
  EXT_ADDRESS_CMD_UNHOLD = 4
  EXT_ADDRESS_CMD_SUSPEND = 5
  EXT_ADDRESS_CMD_UNSUSPEND = 6
  EXT_ADDRESS_CMD_ABORT = 7
  EXT_ADDRESS_CMD_CLEAR = 8
  EXT_ADDRESS_FNC_FREEDRIVE = 9

  global EXT_CtrlCmd = [False, False, False, False, False, False, False, False, False, False]

  EXT_Control_by = "uGO"

  global CMD_Abort = False
  global CMD_Clear = False
  global CMD_Stop = False
  global CMD_Reset = False
  global CMD_Start = False
  global CMD_Hold = False
  global CMD_Unhold = False
  global CMD_Suspend = False
  global CMD_Unsuspend = False
  global FNC_Freedrive = False

  CND_Suspend = False         # condition for suspend command
  CND_Unsuspend = False       # condition for unsuspend command

  thread Get_Pml_Command():
      while (True):
          if (EXT_Control_by == "uGO"):
              EXT_CtrlCmd = ugo_event_controller()
          elif (EXT_Control_by == "Leitsystem"):
              # EXT_CtrlCmd = Leitsystem
          end
          # ---------- Abort ---------- #
          if ((not STATE == 15) and (not STATE == 16) and EXT_CtrlCmd[EXT_ADDRESS_CMD_ABORT]):
              CMD_Abort = True
              CMD_Stop = False
          elif ((STATE == 17) and not EXT_CtrlCmd[EXT_ADDRESS_CMD_ABORT]):
              CMD_Abort = False
          end
          # ---------- Stop ---------- #
          if ((not STATE == 1) and (not STATE == 2) and (get_standard_digital_in(IO_ADDRESS_CMD_STOP) or EXT_CtrlCmd[EXT_ADDRESS_CMD_STOP])):
              CMD_Stop = True
              if get_standard_digital_in(IO_ADDRESS_CMD_STOP):
                  log_state("Stop command by pushbutton")
              elif EXT_CtrlCmd[EXT_ADDRESS_CMD_STOP]:
                  log_state("Stop command by external control")
              end
          elif (STATE == 2) and (not get_standard_digital_in(IO_ADDRESS_CMD_STOP)) and (not EXT_CtrlCmd[EXT_ADDRESS_CMD_STOP]):
              CMD_Stop = False
          end
          CMD_Hold = (STATE == 6 or STATE == 10) and not CMD_Stop and (ERROR.FLAG or EXT_CtrlCmd[EXT_ADDRESS_CMD_HOLD])
          CMD_Reset = (STATE == 2 or STATE == 8) and not CMD_Stop and (read_input_boolean_register(5) or EXT_CtrlCmd[EXT_ADDRESS_CMD_RESET])
          CMD_Start = (STATE == 4) and not CMD_Stop and (get_standard_digital_in(IO_ADDRESS_CMD_START) or EXT_CtrlCmd[EXT_ADDRESS_CMD_START])
          CMD_Unhold = (STATE == 10) and not CMD_Stop and (get_standard_digital_in(IO_ADDRESS_CMD_START) or EXT_CtrlCmd[EXT_ADDRESS_CMD_UNHOLD])
          CMD_Suspend = (STATE == 6) and not CMD_Stop and (CND_Suspend or EXT_CtrlCmd[EXT_ADDRESS_CMD_SUSPEND])
          CMD_Unsuspend = (STATE == 13) and not CMD_Stop and (CND_Unsuspend or EXT_CtrlCmd[EXT_ADDRESS_CMD_UNSUSPEND])
          CMD_Clear = (STATE == 16) and EXT_CtrlCmd[EXT_ADDRESS_CMD_CLEAR]
          FNC_Freedrive = (STATE == 10) and EXT_CtrlCmd[EXT_ADDRESS_FNC_FREEDRIVE]
          sleep(0.1)
      end
  end

  thread_pml_command_handler = run Get_Pml_Command()

  def command_manager(external_control="uGO", cond_suspend=False, cond_unsuspend=False):

      EXT_Control_by = external_control
      CND_Suspend = cond_suspend
      CND_Unsuspend = cond_unsuspend

      if (CMD_Abort and STATE != 15 and STATE != 16):
          STATE = 15
      elif (CMD_Stop and STATE != 1 and STATE != 2):
          STATE = 1
      end
      return False
  end

  def stopping():
      if (EXT_Control_by == "uGO"):
          return ugo_pml_stopping()
      elif (EXT_Control_by == "Leitsystem"):
          # EXT_CtrlCmd = Leitsystem
      else:
          return True
      end
      return False
  end

  def resetting():
      if (EXT_Control_by == "uGO"):
          return ugo_pml_resetting()
      elif (EXT_Control_by == "Leitsystem"):
          # EXT_CtrlCmd = Leitsystem
      else:
          return True
      end
      return False
  end

  def starting():
      if (EXT_Control_by == "uGO"):
          return ugo_pml_starting()
      elif (EXT_Control_by == "Leitsystem"):
          # EXT_CtrlCmd = Leitsystem
      else:
          return True
      end
      return False
  end

  def holding():
      if (EXT_Control_by == "uGO"):
          return ugo_pml_holding()
      elif (EXT_Control_by == "Leitsystem"):
          # EXT_CtrlCmd = Leitsystem
      else:
          return True
      end
      return False
  end

  def unholding():
      if (EXT_Control_by == "uGO"):
          return ugo_pml_unholding()
      elif (EXT_Control_by == "Leitsystem"):
          # EXT_CtrlCmd = Leitsystem
      else:
          return True
      end
      return False
  end

  def suspending():
      if (EXT_Control_by == "uGO"):
          return ugo_pml_suspending()
      elif (EXT_Control_by == "Leitsystem"):
          # EXT_CtrlCmd = Leitsystem
      else:
          return True
      end
      return False
  end

  def unsuspending():
      if (EXT_Control_by == "uGO"):
          return ugo_pml_unsuspending()
      elif (EXT_Control_by == "Leitsystem"):
          # EXT_CtrlCmd = Leitsystem
      else:
          return True
      end
      return False
  end

  def completing():
      if (EXT_Control_by == "uGO"):
          return ugo_pml_completing()
      elif (EXT_Control_by == "Leitsystem"):
          # EXT_CtrlCmd = Leitsystem
      else:
          return True
      end
      return False
  end

  def aborting():
      if (EXT_Control_by == "uGO"):
          return ugo_pml_aborting()
      elif (EXT_Control_by == "Leitsystem"):
          # EXT_CtrlCmd = Leitsystem
      else:
          return True
      end
      return False
  end

  def clearing():
      if (EXT_Control_by == "uGO"):
          return ugo_pml_clearing()
      elif (EXT_Control_by == "Leitsystem"):
          # EXT_CtrlCmd = Leitsystem
      else:
          return True
      end
      return False
  end
  $ 8 "Script: SCRIPT Utility V5.5.script"
  #*****************************************************
  # customer          :   tbd
  # project name      :   tbd
  #****************************************************
  # controller        :
  # software          :
  #****************************************************
  # author            :   P. Koehnke (+49 1628859904; p.koehnke@unitedrobotics.group)
  # Copyright (c)     :   United Robotics Group Health and Food GmbH
  #                       An der Riede 2
  #                       28816 Stuhr
  #                       Germany
  #****************************************************
  # description       :   utility programs for the application
  # version:      	:   3.1
  # created           :   30.01.2023
  # updated           :
  #****************************************************
  # modifications     :   get_tool_free_pose_2(), get_index_from_list()
  #
  # date              :   05.01.2024
  # name              :   PK
  # reason            :
  #****************************************************

  def found_in_matrix(data, req_id, req_idx):
      local id = -1
      local dimensions = size(data)
      local loop_dataset = 0

      while (id != req_id and loop_dataset < dimensions[0]):
          id = data[loop_dataset, 0]
          if (id == req_id):
              return data[loop_dataset, req_idx]
          else:
              loop_dataset = loop_dataset + 1
          end
      end
  end

  def found_in_list(value, list):
      local idx = 0

      while (idx < length(list)):
          if (value == list[idx]):
              return True
          end
          idx = idx + 1
      end
      return False
  end

  def get_index_from_list(list, value = -1):
      local idx = 0

      while (idx < length(list)):
          if (value == -1):
              if (list[idx] != 0):
                  return idx
              end
          else:
              if (list[idx] == value):
                  return idx
              end
          end
          idx = idx + 1
      end
      return -1
  end

  def find_object_by_type(list, type=0):
      local object = list[0]
      local i = 0

      while i < length(list):
          object = list[i]
          if object.type == type:
              return object
          end
          i = i + 1
      end
  end

  def pose_RPY2RotVec(pose):
      local rotvec = rpy2rotvec([d2r(pose[3]), d2r(pose[4]), d2r(pose[5])])
      return p[pose[0], pose[1], pose[2], rotvec[0], rotvec[1], rotvec[2]]
  end

  def pose_RotVec2RPY(pose):
      local rpy = rotvec2rpy([pose[3], pose[4], pose[5]])
      return p[pose[0], pose[1], pose[2], r2d(rpy[0]), r2d(rpy[1]), r2d(rpy[2])]
  end

  def swivel(frame_ref, angles = [0, 0, 0], pose = p[0, 0, 0, 0, 0, 0]):

      local rpy_ref = [0, 0, 0]
      local rpy_new = [0, 0, 0]
      local rotvec_new = [0, 0, 0]
      local pose_from = p[0, 0, 0, 0, 0, 0]
      local pose_to = p[0, 0, 0, 0, 0, 0]
      local i = 0

      if (pose == p[0, 0, 0, 0, 0, 0]):
          pose_to = pose_trans(pose_inv(frame_ref), get_actual_tcp_pose())
      else:
          pose_to = pose
      end

      rpy_ref = rotvec2rpy(frame_ref[3], frame_ref[4], frame_ref[5])

      while (i < 3):
          rpy_new[i] = rpy_ref[i] + d2r(angles[i])
          i = i + 1
      end

      rotvec_new = rpy2rotvec(rpy_new)
      pose_from = p[0, 0, 0, rotvec_new[0], rotvec_new[1], rotvec_new[2]]
      pose_to = p[pose_to[0], pose_to[1], pose_to[2], rotvec_new[0], rotvec_new[1], rotvec_new[2]]

      return pose_trans(pose_from, pose_to)
  end

  def get_random_pose(pose_ref, mode = "", range_max = [0, 0, 0]):
      # modi: "cubic", "rotation"
      # getting a random pose in the x/y-plane. range can be set for each
      # translation and rotation.
      local rpy_random = [0, 0, 0]
      local rotvec_random = [0, 0, 0]
      local pose_random = pose_ref
      local i = 0

      if (mode == "cubic"):
          # cubic mode: random pose takes only x, y and z
          i = 0
          while (i < 3):
              pose_random[i] = pose_ref[i] + range_max[i] * (random() - 0.5)
              i = i + 1
          end
          return pose_random

      elif (mode == "rotation"):
          i = 0
          while (i < 3):
              rpy_random[i] = d2r(range_max[i]) * (random() - 0.5)
              i = i + 1
          end
          rotvec_random = rpy2rotvec(rpy_random)
          pose_random = pose_trans(p[0, 0, 0, rotvec_random[0], rotvec_random[1], rotvec_random[2]], pose_ref)
          return pose_random

      else:
          # unknown mode, return pose_ref
          return pose_ref
      end
  end

  def get_pattern_pos_rectangle(counter, direction, pattern, patterninc = [0, 0], patternsize = [0, 0]):
      # defines the position inside a rectangular pattern
      # pattern describes, how many objects are in x-direction and how many in y-direction [x, y]
      # patternsize will give the total length of each direction [x, y]
      local X_Fac = 0
      local Y_Fac = 0
      local max = pattern[0] * pattern[1]
      local i = 0

      if (1 > counter or counter > max):
          counter = 1
      end

      if pattern[0] == 0:
          pattern[0] = 1
      end

      if pattern[1] == 0:
          pattern[1] = 1
      end

      if (direction == "Y" or direction == "y"):
          X_Fac = floor((counter - 1) / pattern[1])
          Y_Fac = (counter - 1) % pattern[1]
      elif (direction == "X" or direction == "x"):
          X_Fac = (counter - 1) % pattern[0]
          Y_Fac = floor((counter - 1) / pattern[0])
      end

      if patternsize != [0, 0]:
          while i < 2:
              if pattern[i] > 1:
                  patterninc[i] = patternsize[i] / (pattern[i] - 1)
              end
              i = i + 1
          end
      end

      return p[X_Fac * patterninc[0], Y_Fac * patterninc[1], 0, 0, 0, 0]
  end

  def get_pattern_pos_circle(counter, radius, angle, direction, pattern, patternsize = [0, 0]):
      # get the patternpos for a circular pattern through a counter
      # need the radius and the angle in radiants
      local X_Fac = 0
      local Y_Fac = 0
      local rad_bow = 0
      local radius_cal = 0
      local ref = p[0, 0, 0, 0, 0, 0]

      if pattern[0] == 0:
          pattern[0] = 1
      end

      if pattern[1] == 0:
          pattern[1] = 1
      end

      if (direction == "Y" or direction == "y"):
          X_Fac = floor((counter - 1) / pattern[1])
          Y_Fac = (counter - 1) % pattern[1]
      elif (direction == "X" or direction == "x"):
          X_Fac = (counter - 1) % pattern[0]
          Y_Fac = floor((counter - 1) / pattern[0])
      end

      # the opening angle will be calculated in x-direction
      # works only between -90 and 90 degree
      if pattern[0] > 1:
          rad_bow = - angle / (pattern[0] - 1) * X_Fac + angle / 2
      end

      if (counter % 2 == 0 and pattern[1] > 1):
          radius_cal = radius - patternsize[1] / (pattern[1])
      else:
          radius_cal = radius + patternsize[1] / (pattern[1])
      end
      ref = p[0, radius_cal, 0, 0, 0, 0]

      return p[ref[0] * cos(rad_bow) - ref[1] * sin(rad_bow), (ref[0] * sin(rad_bow) + ref[1] * cos(rad_bow)) - radius, 0, 0, 0, 0]
  end

  def get_pattern_counter(pose, direction, pattern, patterninc = [0, 0], patternsize = [0, 0]):
      # returns the counter for a pattern from a given cartesian pose
      local patternpose = p[pose[0], pose[1], 0, 0, 0, 0]
      local X_Fac = 0
      local Y_Fac = 0
      local i = 0

      if patternsize != [0, 0]:
          while i < 2:
              if pattern[i] > 1:
                  patterninc[i] = patternsize[i] / (pattern[i] - 1)
              else:
                  pattern[i] = 0
              end
              i = i + 1
          end
      end

      # calculation of the counter in the desired axis-direction
      if (direction == "x" or direction == "X"):
          if patterninc[0] > 0:
              X_Fac = ceil((patternpose[0] + patterninc[0] / 2) / patterninc[0])
              if X_Fac < 0:
                  X_Fac = 0
              end
          end
          if patterninc[1] > 0:
              Y_Fac = floor((patternpose[1] + patterninc[1] / 2) / patterninc[1])
              if Y_Fac < 0:
                  Y_Fac = 0
            end
          end
          return Y_Fac * pattern[0] + X_Fac
      elif (direction == "y" or direction == "Y"):
          if patterninc[0] > 0:
              X_Fac = floor((patternpose[0] + patterninc[0] / 2) / patterninc[0])
          end
          if patterninc[1] > 0:
              Y_Fac = ceil((patternpose[1] + patterninc[1] / 2) / patterninc[1])
          end
          return X_Fac * pattern[1] + Y_Fac
      end
  end

  def get_plc_reg(mod_sig_name):
      return integer_to_binary_list(modbus_get_signal_status(mod_sig_name))
  end

  def set_plc_reg(mod_sig_name, mod_sig_list):
      modbus_set_output_register(mod_sig_name, binary_list_to_integer(mod_sig_list), False)
  end

